(* IEC 61131-3 sources: daoli-st-library/DL_Motion (part 24) *)

(* ---- FB_DL_MotionCmdQueue.st ---- *)
(*
    FB_DL_MotionCmdQueue —— 运动指令排队器（仅 Buffered 语义）
    ------------------------------------------------------------------
    分类      : DL_Motion / CommandMgmt
    前缀      : FB_DL_
    版本      : 1.0.1
    溯源      : T1-6 PLCopen MC_BUFFERMODE 公开条款（Aborting / Buffered / BlendingLow /
                BlendingHigh / BlendingPrevious / BlendingNext 六种，其中 Buffered
                = 「新指令等前一条 Done 之后才影响轴」）；本件只实现 Buffered 一种；
                环形缓冲、满队策略、去重、自愈规则与码位 100% 自有；clean-room 重写，
                未复制任何闭源厂商源码，参考实现仅限 MIT/Apache 许可
    道莅 clean-room 防御性实现：语义借鉴、代码与码位 100% 自有
    平台      : 纯 IEC 61131-3，CODESYS V3.5+ / TwinCAT 3 / InoProShop / Machine Expert 通用
    作者      : 道莅代码库 · PLC编程专家（R22 批 4 · #14）
    ------------------------------------------------------------------
    功能说明  : 把上位连发的定位指令排成先入先出队列，按 Buffered 语义一条一条放给轴：
                前一条轴的 Done 未回就不发下一条。本件不消费轴状态、不发 MC_ 功能块、
                不判断运动是否成功——轴的 Done / Error 由调用方以引脚注入。
    职责边界  : ① 只做 Buffered。Blending 系列不立：BlendingLow / BlendingHigh /
                   BlendingPrevious / BlendingNext 都要求「两段速度在过渡点融合」，
                   而本库的轴侧接口没有速度融合通道，硬做只能做出假混合，
                   比不做更危险——故明确不立项，调用方需融合时请用轴厂家的原生接口。
                ② 不做指令合法性（软限位、速度上限）判定，那是 FB_DL_SoftLimitGuard 的职责。
                ③ bAxisError 到达后只挂起不自动续发：必须先让轴故障消失、再给 bClear，
                   否则队列会在轴仍故障时继续往下砸指令，那是二次伤害。
    队列实现  : 环形缓冲，深度固定 DL_MQ_DEPTH = 8（不参数化：动态内存违反零厂商依赖）。
                头指针指向待发条目，尾指针指向下一个空位，计数 _uCount 为权威值。
    自愈规则  : 每拍前置一致性检查，规则写在此处即此件的契约：
                ① 头指针、尾指针任一 >= DL_MQ_DEPTH，或计数 > DL_MQ_DEPTH
                   → 指针与内容均不可信，整队重建（计数与双指针全部归零）；
                ② 指针均合法时，用 (尾 − 头 + 深度) MOD 深度 反算应有计数，
                   满队时该值为 0，按满队解释为 DL_MQ_DEPTH；
                   反算值与 _uCount 不符 → 以指针为准重建计数（双指针是同拍维护的，
                   计数可能被外部复位或掉电字节残留破坏，指针更可信）。
                自愈是静默的，不占码位（不影响工艺判定），但会在头注释留档供现场排查。
    偏离留档  : 派单写「bAxisDone 上升沿出队」，若按字面在 Done 那一拍才移出队首，
                bClear 期间的槽位归属会与新入队条目混叠（新条目可能被下一次 Done 误当成
                在飞条目弹出，等于吞掉一条指令）。本件把「出队」放在发令那一拍完成，
                Done 只负责把状态机送回 eIdle——语义等价，且消除了混叠路径。
    错误码    : 16#0004_01D9 队列满：bOverwriteOldest=TRUE 丢最旧 / FALSE 拒绝新入队
                              （两策略共用本码，靠 uDropped 是否自增区分）——信息级
                16#0004_01DA 连续同目标同速度的指令已合并去重——信息级，正常防御
                16#0004_02F0 指令参数非有限（NaN / ±Inf），拒绝入队且不占槽——故障级，
                             只拒这一条，不打断整队，也不改变状态机（非锁存）
                16#0004_02F1 轴故障应答（bAxisError），已清队并挂起，禁止自动续发——故障级
                16#0004_02F2 状态机落 ELSE 兜底（非法状态）——故障级，回 eIdle 并清队
    码位总账  : 16#0004_01D9 用 / 16#0004_01DA 用 ｜ 16#0004_02F0 用 / 16#0004_02F1 用 / 16#0004_02F2 用
    状态机    : E_DL_CmdQueueState（eIdle / eSending / eWaitDone / eFault），
                CASE 含 ELSE 兜底，ELSE 置 16#0004_02F2 并回 eIdle 同时清队；
                eSending 是单拍相（发令拍），进相即出相，bExec 因此天然只亮一拍。
    采样约定  : 三个 R_TRIG（入队 / 轴 Done / 轴 Error）在本体最前部无条件刷新（R40）；
                bExec 由段 2 的预置清零保证单拍（R25 三律：置位后本拍即被预置覆盖，
                下一拍必为 FALSE，不存在只置不清）。
    依赖      : 仅 Standard.library（R_TRIG / ABS / MIN / MAX），不引用任何其他 DL_ 子库。
    验收向量  :
                V1 域外早退：fTargetPos = NaN 入队 → 02F0、bError=TRUE、uCount 不变、
                   不占槽，整队继续可用。
                V2 上限截断：连发 9 条 → 第 9 条时 bFull=TRUE；bOverwriteOldest=TRUE
                   → uDropped=1、uCount 仍 8、01D9；置 FALSE → uDropped 不变、01D9、
                   新条目被拒。
                V3 跨段时序：eWaitDone 中 bAxisDone 与下一次 bEnq 同拍 → 本拍先入队
                   （uCount+1）再出相；下一拍才发令，bExec 不连拍。
                V4 恢复首拍：bAxisError 上升沿 → 02F1、清队、eFault；轴故障消失后
                   单独给 bClear → 回 eIdle，队列为空且不发任何残留指令。
    红线自检  : 1 全局变量声明零使用 / 外部变量访问零使用 / 物理地址零使用 —— 通过，全部量经引脚注入
                2 纯 IEC 61131-3 跨平台 —— 通过，仅 Standard.library，无动态内存
                3 防御性编程 —— 通过，数组索引全部前置界检、计数递减前判零、
                   浮点判等用 1.0E-6 容差、非有限值拒绝入队
                4 声明行同行中英双语注释 + 单位 —— 通过，逐行附注（含枚举与数组）
                5 ENUM + CASE 且含 ELSE 兜底 —— 通过
                6 TON / R_TRIG 无条件刷新 —— 通过，段 1 三个沿实例先行调用
                7 无魔法数 —— 通过，深度、容差、计数上限全部 VAR CONSTANT
    修订记录  : 2026-11-16 v1.0.0 首次入库（R22 批 4 · #14）
                2026-11-16 v1.0.1 R22 终审修复：eSending 进相后队列若被 bClear /
                轴故障清空，发令被跳过时改回 eIdle，不再空等永不到来的轴 Done
                （消除「清队竞态 → eWaitDone 挂死」路径，新增 V5 验收向量：
                eIdle 转 eSending 的下一拍给 bClear → 本拍不发令、回 eIdle、bExec 不出现）
*)
TYPE E_DL_CmdQueueState :
(
    eIdle     := 0,      // 空闲，队列非空即进发令相 / idle, a non-empty queue enters the sending phase
    eSending  := 10,     // 单拍发令相，本拍出队并把指令放到执行引脚 / one-scan sending phase, dequeues and publishes the command
    eWaitDone := 20,     // 等轴 Done，未回不发下一条（Buffered 契约）/ waiting for the axis Done, nothing else is issued before it
    eFault    := 30      // 故障，队列已清，需轴故障消失后再给 bClear / fault, the queue is cleared and a bClear is required after the axis fault disappears
);
END_TYPE

FUNCTION_BLOCK FB_DL_MotionCmdQueue
VAR_INPUT
    bEnq             : BOOL;                   // 入队请求，上升沿生效 / enqueue request, effective on the rising edge
    fTargetPos       : REAL;                   // 目标位置 [mm]，非有限即拒收 / target position [mm], a non-finite value is rejected
    fVelocity        : REAL;                   // 运行速度 [mm/s]，非有限即拒收 / travel velocity [mm/s], a non-finite value is rejected
    bAxisDone        : BOOL;                   // 轴 Done 输入，由调用方注入，本件不消费轴状态 / axis Done injected by the caller, no axis state is consumed here
    bAxisError       : BOOL;                   // 轴故障输入，上升沿清队挂起 / axis error input, a rising edge clears the queue and suspends
    bOverwriteOldest : BOOL := TRUE;           // 满队策略：TRUE 丢最旧 / FALSE 拒绝新入队 / full-queue policy, TRUE drops the oldest, FALSE rejects the newcomer
    bClear           : BOOL;                   // 清队电平，为真期间队列保持空且不发令 / clear level, the queue stays empty and nothing is issued while TRUE
END_VAR
VAR_OUTPUT
    bExec            : BOOL;                   // 发令单拍脉冲，只亮一拍 / issue pulse, asserted for exactly one scan
    fExecPos         : REAL;                   // 本拍发出的目标位置 [mm]，保持到下一次发令 / target position issued this scan [mm], held until the next issue
    fExecVel         : REAL;                   // 本拍发出的运行速度 [mm/s]，保持到下一次发令 / travel velocity issued this scan [mm/s], held until the next issue
    uCount           : UINT;                   // 队列内条目数 [条]，0~DL_MQ_DEPTH / number of queued items [pcs], 0~DL_MQ_DEPTH
    bFull            : BOOL;                   // 队列已满 / the queue is full
    uDropped         : UDINT;                  // 累计丢弃条数 [条]，饱和不回绕 / accumulated dropped items [pcs], saturating and never wrapping
    eErr             : UDINT;                  // 错误码，0 表示无错 / error code, 0 means no error
    bError           : BOOL;                   // 故障级标志，仅故障级错误置位 / fault-class flag, set only on fault-level codes
    bValid           : BOOL;                   // 输出可用标志，= NOT bError / outputs valid flag, equals NOT bError
END_VAR
VAR
    fbEnq            : R_TRIG;                 // 入队沿检测实例，无条件刷新 / enqueue edge instance, refreshed unconditionally
    fbDone           : R_TRIG;                 // 轴 Done 沿检测实例，无条件刷新 / axis Done edge instance, refreshed unconditionally
    fbAxisErr        : R_TRIG;                 // 轴故障沿检测实例，无条件刷新 / axis error edge instance, refreshed unconditionally
    _afPos           : ARRAY[0..DL_MQ_DEPTH - 1] OF REAL;   // 队列位置缓存 [mm]，深度与 DL_MQ_DEPTH 同源 / queued positions [mm], depth tied to DL_MQ_DEPTH
    _afVel           : ARRAY[0..DL_MQ_DEPTH - 1] OF REAL;   // 队列速度缓存 [mm/s] / queued velocities [mm/s]
    _uHead           : UINT;                   // 头指针，指向待发条目 / head pointer, points at the next item to issue
    _uTail           : UINT;                   // 尾指针，指向下一个空位 / tail pointer, points at the next free slot
    _uCount          : UINT;                   // 队列条目数（权威值）[条] / item count, the authoritative value [pcs]
    _uExp            : UINT;                   // 由双指针反算的应有计数，自愈用 [条] / count derived from the pointers, used by the self-healing path [pcs]
    _uDroppedAcc     : UDINT;                  // 丢弃计数累加器，饱和不回绕 [条] / dropped accumulator, saturating and never wrapping [pcs]
    _fLastPos        : REAL;                   // 最近一次入队或发令的目标位置，去重用 [mm] / last queued or issued target, used for de-duplication [mm]
    _fLastVel        : REAL;                   // 最近一次入队或发令的速度，去重用 [mm/s] / last queued or issued velocity, used for de-duplication [mm/s]
    _bHaveLast       : BOOL;                   // 去重基准是否已建立 / whether the de-duplication reference exists
    _bParamBad       : BOOL;                   // 本条指令参数非有限标志 / the incoming command carries a non-finite value
    _eState          : E_DL_CmdQueueState;     // 当前状态 / current state
END_VAR
VAR CONSTANT
    DL_MQ_DEPTH      : UINT := 8;              // 队列深度 [条]，固定不参数化 / queue depth [pcs], fixed and never parameterised
    DL_MQ_UDINT_MAX  : UDINT := 16#FFFF_FFFF;  // 丢弃计数饱和上限 [条] / drop-counter saturation bound [pcs]
    DL_MQ_EPS        : REAL := 1.0E-6;         // 去重浮点判等容差 [mm] / de-duplication tolerance [mm]
    DL_MQ_INF_GUARD  : REAL := 4.0E38;         // 非有限幅值判定阈（大于 REAL 最大值）[mm] / non-finite magnitude guard [mm]
END_VAR

// 段 1｜三个沿检测实例无条件周期刷新（红线 6：严禁放入 IF / CASE）
// segment 1, three edge instances refreshed unconditionally
fbEnq(CLK := bEnq);
fbDone(CLK := bAxisDone);
fbAxisErr(CLK := bAxisError);

// 段 2｜输出与错误状态预置（bExec 的单拍性由这里的预置保证，R25 三律）
// segment 2, preset outputs and error status; the preset here is what makes bExec a true one-scan pulse
eErr := 0;                                      // 预置无错误 / preset no error
bError := FALSE;                                // 预置无故障标志 / preset no error flag
bExec := FALSE;                                 // 预置无发令，任何状态想发令必须在本拍重新置位 / preset no issue, any state must assert it again this scan
_bParamBad := FALSE;                            // 预置入队参数合法 / preset the incoming command as legal

// 段 3｜队列自愈：指针越界即整队重建，计数与指针推算不符以指针为准（规则见头注释）
// segment 3, queue self-healing; an out-of-range pointer rebuilds the whole queue and a count mismatch follows the pointers
IF (_uHead >= DL_MQ_DEPTH) OR (_uTail >= DL_MQ_DEPTH) OR (_uCount > DL_MQ_DEPTH) THEN
    _uHead := 0;                                // 指针越界，头归零 / out-of-range head reset
    _uTail := 0;                                // 指针越界，尾归零 / out-of-range tail reset
    _uCount := 0;                               // 内容不可信，计数归零 / untrustworthy content, count reset
    _bHaveLast := FALSE;                        // 去重基准随队一起作废 / the de-duplication reference dies with the queue
ELSE
    _uExp := (_uTail + DL_MQ_DEPTH - _uHead) MOD DL_MQ_DEPTH;   // 由双指针反算应有计数 / derive the count from the pointers
    IF (_uCount > 0) AND (_uExp = 0) THEN
        _uExp := DL_MQ_DEPTH;                   // 满队时头尾重合，按满队解释 / a full queue has coincident pointers, read it as full
    END_IF
    IF _uCount <> _uExp THEN
        _uCount := _uExp;                       // 计数与指针不符，以指针为准重建 / a mismatch follows the pointers, which are maintained every scan
    END_IF
END_IF

// 段 4｜清队电平：只清队列内容，不打断在飞指令的完成等待（Buffered 契约）
// segment 4, the clear level empties the queue but never interrupts the wait of the in-flight command
IF bClear THEN
    _uHead := 0;                                // 头归零 / head reset
    _uTail := 0;                                // 尾归零 / tail reset
    _uCount := 0;                               // 计数归零 / count reset
    _bHaveLast := FALSE;                        // 去重基准作废 / the de-duplication reference is void
END_IF

// 段 5｜轴故障应答：上升沿清队并挂起，绝不自动续发（批 4 统一口径）
// segment 5, axis error response, a rising edge clears the queue and suspends, never resuming automatically
IF fbAxisErr.Q THEN
    _uHead := 0;                                // 头归零 / head reset
    _uTail := 0;                                // 尾归零 / tail reset
    _uCount := 0;                               // 清队，故障后不得留残留指令 / clear the queue, no residual command may survive a fault
    _bHaveLast := FALSE;                        // 去重基准作废 / the de-duplication reference is void
    eErr := 16#0004_02F1;                       // 故障级：轴故障应答已清队并挂起 / fault: the axis error response cleared the queue and suspended
    bError := TRUE;                             // 置故障标志 / raise the fault flag
    _eState := E_DL_CmdQueueState.eFault;       // 挂起，等轴故障消失后再给 bClear / suspend until the axis fault is gone and a bClear arrives
END_IF

// 段 6｜入队处理：参数门禁 → 去重 → 满队策略 → 落槽
// segment 6, enqueue path, parameter gate then de-duplication then the full-queue policy then the slot write
IF fbEnq.Q AND (NOT bClear) AND (_eState <> E_DL_CmdQueueState.eFault) THEN
    // 6.1 参数门禁：非有限一律拒收，不占槽、不动计数
    // parameter gate, a non-finite value is rejected without taking a slot or touching the count
    IF (fTargetPos - fTargetPos) <> (fTargetPos - fTargetPos) THEN
        _bParamBad := TRUE;                     // 目标位置为 NaN / the target position is NaN
    ELSIF ABS(fTargetPos) > DL_MQ_INF_GUARD THEN
        _bParamBad := TRUE;                     // 目标位置为 ±Inf / the target position is infinite
    ELSIF (fVelocity - fVelocity) <> (fVelocity - fVelocity) THEN
        _bParamBad := TRUE;                     // 速度为 NaN / the velocity is NaN
    ELSIF ABS(fVelocity) > DL_MQ_INF_GUARD THEN
        _bParamBad := TRUE;                     // 速度为 ±Inf / the velocity is infinite
    END_IF

    IF _bParamBad THEN
        eErr := 16#0004_02F0;                   // 故障级：指令参数非有限，拒收 / fault: non-finite command parameter, rejected
        bError := TRUE;                         // 只拒这一条，不打断整队 / rejects this item only and never disturbs the rest of the queue
    ELSIF _bHaveLast
          AND (ABS(fTargetPos - _fLastPos) <= DL_MQ_EPS)
          AND (ABS(fVelocity - _fLastVel) <= DL_MQ_EPS) THEN
        eErr := 16#0004_01DA;                   // 信息级：与最近一条同目标同速度，合并去重 / info: identical to the latest command, merged
    ELSIF _uCount >= DL_MQ_DEPTH THEN
        // 6.2 满队：按策略处理，两种策略共用 01D9，靠 uDropped 是否自增区分（R90）
        // full queue, both policies share 01D9 and are told apart by whether uDropped grows
        IF bOverwriteOldest AND (_uCount > 0) THEN
            _uHead := (_uHead + 1) MOD DL_MQ_DEPTH;     // 丢最旧：头前移一格 / drop the oldest by advancing the head
            _uCount := _uCount - 1;                     // 计数先减，随后落槽再加回 / decrement first, the slot write adds it back
            IF _uDroppedAcc < DL_MQ_UDINT_MAX THEN
                _uDroppedAcc := _uDroppedAcc + 1;       // 丢弃计数饱和自增 / saturating increment of the drop counter
            END_IF
            _afPos[_uTail] := fTargetPos;               // 落槽（索引已由指针范围检查保证合法）/ write the slot, the index was validated by the pointer check
            _afVel[_uTail] := fVelocity;                // 落槽速度 / write the queued velocity
            _uTail := (_uTail + 1) MOD DL_MQ_DEPTH;     // 尾前移一格 / advance the tail
            _uCount := _uCount + 1;                     // 计数加回 / add the count back
            _fLastPos := fTargetPos;                    // 更新去重基准位置 / update the de-duplication reference
            _fLastVel := fVelocity;                     // 更新去重基准速度 / update the de-duplication reference
            _bHaveLast := TRUE;                         // 基准已建立 / the reference now exists
            eErr := 16#0004_01D9;                       // 信息级：队列满，已丢最旧 / info: the queue was full and the oldest was dropped
        ELSE
            eErr := 16#0004_01D9;                       // 信息级：队列满，拒绝新入队（uDropped 不变）/ info: full and the newcomer is rejected, uDropped stays
        END_IF
    ELSE
        _afPos[_uTail] := fTargetPos;           // 落槽（索引已由指针范围检查保证合法）/ write the slot, the index was validated by the pointer check
        _afVel[_uTail] := fVelocity;            // 落槽速度 / write the queued velocity
        _uTail := (_uTail + 1) MOD DL_MQ_DEPTH; // 尾前移一格 / advance the tail
        _uCount := _uCount + 1;                 // 计数加一 / increment the count
        _fLastPos := fTargetPos;                // 更新去重基准位置 / update the de-duplication reference
        _fLastVel := fVelocity;                 // 更新去重基准速度 / update the de-duplication reference
        _bHaveLast := TRUE;                     // 基准已建立 / the reference now exists
    END_IF
END_IF

// 段 7｜状态机：eIdle 取队首 → eSending 单拍发令并出队 → eWaitDone 等 Done → eIdle
// segment 7, the state machine, take the head in eIdle, issue and dequeue in the one-scan eSending phase, then wait for Done
CASE _eState OF
E_DL_CmdQueueState.eIdle:
    IF (_uCount > 0) AND (NOT bClear) THEN
        _eState := E_DL_CmdQueueState.eSending;     // 有货且未清队，进发令相 / there is work and no clear, enter the sending phase
    END_IF

E_DL_CmdQueueState.eSending:
    IF (_uCount > 0) AND (_uHead < DL_MQ_DEPTH) THEN
        fExecPos := _afPos[_uHead];                 // 读队首位置（索引前置界检）/ read the head position with a bounds check
        fExecVel := _afVel[_uHead];                 // 读队首速度 / read the head velocity
        bExec := TRUE;                              // 单拍发令，段 2 的预置保证下一拍必为 FALSE / the one-scan issue, the preset guarantees FALSE next scan
        _fLastPos := fExecPos;                      // 去重基准同步为已发条目 / the de-duplication reference follows the issued item
        _fLastVel := fExecVel;                      // 去重基准同步为已发条目 / the de-duplication reference follows the issued item
        _bHaveLast := TRUE;                         // 基准已建立 / the reference now exists
        _uHead := (_uHead + 1) MOD DL_MQ_DEPTH;     // 出队在发令这一拍完成，避免与 bClear 混叠 / dequeue right here so bClear cannot alias the slot
        _uCount := _uCount - 1;                     // 上面的 _uCount > 0 判断已挡住无符号下溢 / the guard above prevents an unsigned underflow
        _eState := E_DL_CmdQueueState.eWaitDone;    // 已真实发令：本相转入等待轴 Done / issued for real, now wait for the axis Done
    ELSE
        _eState := E_DL_CmdQueueState.eIdle;        // 进相后队列被 bClear / 故障清空：无在飞指令，直接回空闲，不得空等永不出现的 Done（R22 终审修复：消除竞态挂死）/ the queue was emptied after entering this phase, no command is in flight, return to idle instead of waiting forever
    END_IF

E_DL_CmdQueueState.eWaitDone:
    IF fbDone.Q THEN
        _eState := E_DL_CmdQueueState.eIdle;        // 前条完成，允许发下一条 / the previous move is done and the next may be issued
    END_IF

E_DL_CmdQueueState.eFault:
    // 退出条件：轴故障已消失且人来清队——两者缺一不可，绝不自动续发
    // exit needs both a vanished axis fault and an operator clear, no automatic resume
    IF bClear AND (NOT bAxisError) AND (NOT fbAxisErr.Q) THEN
        _eState := E_DL_CmdQueueState.eIdle;        // 允许回空闲，队列此时已空；进入故障的这一拍不得退出，否则故障码只闪一拍 / back to idle, but never on the entering scan or the fault code would flash for a single scan
    END_IF

ELSE
    eErr := 16#0004_02F2;                           // 故障级：状态机落 ELSE / fault: the state machine fell into ELSE
    bError := TRUE;                                 // 置故障标志 / raise the fault flag
    _uHead := 0;                                    // 非法态一律清队，绝不带着未知队列继续跑 / an illegal state always clears the queue
    _uTail := 0;
    _uCount := 0;
    _bHaveLast := FALSE;                            // 去重基准作废 / the de-duplication reference is void
    _eState := E_DL_CmdQueueState.eIdle;            // 回空闲 / back to idle
END_CASE

// 段 8｜出口汇总：计数类只做发布，不再二次改写（禁隐式回夹）
// segment 8, exit aggregation; counters are published here and never rewritten again
uCount := _uCount;                              // 队列条目数发布 [条] / publish the queued item count [pcs]
uDropped := _uDroppedAcc;                       // 丢弃累计发布 [条] / publish the accumulated drops [pcs]
bFull := (_uCount >= DL_MQ_DEPTH);              // 满队标志 / full-queue flag
bValid := NOT bError;                           // 输出可用 = 无故障级错误 / outputs are valid when no fault-level code is present
END_FUNCTION_BLOCK

(* ---- FB_DL_PassiveHomingMonitor.st ---- *)
(*==============================================================================
 * 组件名称 (Component)  : FB_DL_PassiveHomingMonitor
 * 所属子库 (Sublibrary) : DL_Motion
 * 当前版本 (Version)    : 1.0.1
 * 组件分类 (Category)   : 功能块（FUNCTION_BLOCK）· 被动回零旁路监听（参考事件确认）
 * 兼容性   (Platform)   : CODESYS 3.5 / TwinCAT 3 / 汇川 InoProShop / Schneider Machine Expert
 *                         仅依赖 Standard.library（R_TRIG / F_TRIG / TON / ABS / MIN / MAX / LIMIT）
 * 接口依赖 (Depends)    : 无 DL_ 内部依赖。本件**不引用**轴状态枚举、**不定义**轴状态枚举，
 *                         也**不调用**任何 MC_ 运动功能块（见分层声明）。
 * 功能描述 (Function)   : 轴被外力移动时（手摇轮、另一驱动拖动、重力下落、维护推车），
 *                         旁路监听参考事件（原点开关沿 / Z 相 / 标记锁存），按「方向一致性
 *                         + 速度窗 + 多次位置一致性」三条判据确认参考点，输出建议施加的
 *                         位置偏移给上层，由上层以 MC_SetPosition 语义消费。
 * 边界（最重要）        : **不自造轴状态、不写轴状态机**。本件只有一个工艺位 bReferenced，
 *                         轴状态（Disabled / Standstill / DiscreteMotion 等）**只由运动层
 *                         拥有**——这是 R31 家族（两套状态机并存）的最高危区，本件按 R11
 *                         判例执行：输出相位 ePhase 仅供 HMI 诊断显示，**不得**被上层当作
 *                         轴状态使用，也不得反向改写轴状态位。
 *                         与 FB_DL_AxisHomingSeq 的分工：后者是**主动回零顺控**（自己发运动
 *                         指令、四模式），本件**不发任何运动指令**，只旁路监听并输出偏移；
 *                         两者可并存，但不得互相改写对方的结论位。
 * 分层声明 (Layer)      : 运动层旁路监视件。上行只为「建议偏移」，下行只有引脚采样。
 *                         零全局变量表引用、零外部变量声明、零物理 IO 地址。
 * 段序     (Segments)   : 段1 实例无条件刷新 → 段2 复位通道（CASE 前，R39）→ 段3 撤防受理 →
 *                         段4 输入防御与镜像量锁定 → 段5 布防受理（倒计置位点，R34）→
 *                         段6 事件受理（倒计递减点，与段5 相邻，R34）→ 段7 状态机 →
 *                         段8 码位单一优先级链 → 段9 出口钳位与保持语义重写。
 * 枚举映射表 (R31)      : eIdle(0)→标签 0｜eArmed(10)→标签 10｜eCaptured(20)→标签 20｜
 *                         eConfirmed(30)→标签 30｜eTimeout(40)→标签 40｜eFault(99)→标签 99。
 *                         每个成员有且仅有一个显式标签，ELSE 只接脏值（02D4）。
 * 单拍标志清单 (R25)    : bArm —— 预清零点：段1 每拍由 `_bArmReq := FALSE` 前的实例输出覆盖；
 *                         置位点：段1 `_bArmReq := _fbTrigArm.Q AND (NOT _bArmConsumed)`；
 *                         自清点：段5 消费时 `_bArmConsumed := TRUE`（撤防、超时、复位三处解除）。
 *                         bReset —— 预清零点：段1 每拍覆盖 _bResetEdge；置位点：段1 的
 *                         _fbTrigReset 实例调用；自清点：紧随实例调用的 _bResetEdge 赋值行。
 *                         bRefEvent —— 内部取上升沿（段1 实例），在段6 单点消费，无对外单拍位。
 * 保持位清单 (R27)      : bReferenced / fRefPos / fOffsetToApply —— 三者逐拍由
 *                         _bRefLatched / _fRefPosHeld / _fOffsetHeld 重写并夹域；
 *                         nEventCount 逐拍由 _nEventCount 转换重写。复位沿清结论。
 * 定时器清单 (R40)      : _fbTonArmTimeout｜IN = (相位 = eArmed 或 eCaptured) AND NOT _bArmBreak｜
 *                         断输入标志 _bArmBreak（每次布防置一拍，本拍 TON 复位 ET）｜
 *                         自清点：段3 无条件 `IF _bArmBreak THEN _bArmBreak := FALSE; END_IF`。
 *                         _fbTonNoMotion｜IN = (相位 = eArmed 或 eCaptured) AND NOT bInMotion
 *                         AND NOT _bArmBreak｜语义为「布防期间长时间静止」信息码 01C5。
 * 三元一致表 (R35)      : 速度窗下限守卫 0.01~100 mm/s / 封顶 100 / 判据 `<`（低于即降精度）｜
 *                         速度窗上限守卫 1~10000 mm/s / 封顶 10000 / 判据 `>`（高于即降精度）｜
 *                         一致性容差守卫 0.001~10 mm / 封顶 10 / 判据 `>`（超出即计数重置）。
 * 镜像量清单 (R38)      : fActPos 的唯一消费点是 _fPosSnap（段4 锁定），fActVel 的唯一消费点
 *                         是 _fVelSnap（段4 锁定）；事件受理与限幅判定全部读快照，不读实时入参。
 * 开源溯源 (Origin)     : 原创实现（参考 PLCopen Part 1 的「参考事件（reference event）」与
 *                         被动回零（passive homing）公开语义，T1-6：参考事件上升沿捕获、
 *                         方向一致性、速度窗内采信、多次事件一致性确认，全部为公开的
 *                         技术概念；实现、状态机、码位与引脚契约 100% 本库独立设计，
 *                         clean-room 编写，未复制任何源码行。许可证说明：PLCopen 规范为
 *                         公开规范条款（非代码），引用其条款语义不构成代码复制风险；
 *                         本文件为本库原创，随本库许可证发布。
 * 验收向量 (Acceptance) :
 *   V1 布防 → 正向 20 mm/s → 两次事件（100.00 / 100.05 mm）→ bReferenced = TRUE、
 *      fRefPos = 100.025（取算术均值，非取首个事件，见设计要点③）。
 *   V2（V-C 方向反转）第二次事件发生在反向 → 16#0004_01C4、计数回到 1、**不得**确认。
 *   V3（V-D 超时恢复）tArmTimeout 到 → eTimeout + 16#0004_02D2；重新 bArm 后计数从 0 重建
 *      （R41：恢复不重头，不允许沿用上次部分计数）。
 *   V4（V-A 非有限）fActVel = NaN → 16#0004_02D3、fRefPos 保持上次确认值（不写脏值）。
 *   V5（R43 出口夹域）撤防后 fOffsetToApply 保持上次值且夹进 ±1.0E6 mm；冷启动首拍输出 0.0。
 * 偏离留档 (Deviation)  :
 *   ① 「目标位置」来源：规格要求输出 fOffsetToApply = 目标 − 参考，但引脚表未给目标值引脚。
 *      本件按「参考事件处应读 0.0 mm」的通用约定输出 fOffsetToApply = 0.0 − fRefPos；若现场
 *      参考点非 0，调用方在消费时叠加其目标值（不新增引脚，避免破坏已冻结的引脚契约）。
 *   ② 速度窗上限的处置：规格给 01C3 的语义是「低于窗下限，采信但精度降级」。高于上限时
 *      定位精度同样不保（可能漏捕获相邻事件），本件并入同一信息码 01C3，语义记为「速度窗
 *      越界，已采信但精度降级」，不新增码位（码位表以规格为准）。
 *   ③ fVelMin > fVelMax 时按对调修复并保持静默（无对应码位），属参数自愈，不改变判定逻辑。
 * 修订历史 (Revision)   :
 *   2026-11-15  v1.0.0  首版入库（Round 13 · 泳道 C · DL_Motion 第 18 件，补 R8 留扩产项）
 *   2026-11-16  v1.0.1  终审修复：段6 事件受理条件补串 bEnable 与 NOT _bFaultCond ——
 *                       原实现下，非有限值检出当拍若恰有参考事件沿，零化快照会被采信，
 *                       极端情形把 0.0 锁存为参考点（坏值穿透到 bReferenced 保持位）
 *============================================================================*)

(*-----------------------------------------------------------------------------
 * 枚举: E_DL_PassiveHomePhase（归属 FB_DL_PassiveHomingMonitor，同文件发布）
 * 用途: 仅内部相位与 HMI 诊断显示，**不是**轴状态，禁止被上层当作轴状态使用。
 *----------------------------------------------------------------------------*)
TYPE E_DL_PassiveHomePhase :
(
    eIdle      := 0,    // 空闲：未布防 / Idle, not armed
    eArmed     := 10,   // 已布防：等待首个参考事件 / Armed, awaiting the first reference event
    eCaptured  := 20,   // 已捕获：事件数未达标，等待后续一致性事件 / Captured, awaiting consistent events
    eConfirmed := 30,   // 已确认：参考点成立，结论保持 / Confirmed, reference established and held
    eTimeout   := 40,   // 超时：布防期内未捕获足够事件 / Timeout, not enough events while armed
    eFault     := 99    // 故障：位置或速度非有限 / Fault, non-finite position or velocity
) UINT;
END_TYPE

FUNCTION_BLOCK FB_DL_PassiveHomingMonitor
VAR_INPUT
    bEnable          : BOOL;                // 使能（Enable），FALSE = 冻结监听并清布防；复位通道不受其屏蔽 / Enable, FALSE stops monitoring
    bReset           : BOOL;                // 复位（Reset），上升沿清结论与锁存 / Rising edge clears the verdict and latches
    bArm             : BOOL;                // 布防（Arm），上升沿开始监听，下降沿撤防 / Rising edge arms, falling edge disarms
    bRefEvent        : BOOL;                // 参考事件电平（Raw reference event），内部取上升沿 / Raw reference event, edge detected inside
    bDirForward      : BOOL := TRUE;        // 本拍运动方向（Current direction），TRUE = 正向，默认 TRUE / TRUE forward, FALSE reverse
    fActPos          : REAL;                // 实际位置（Actual position）[mm]，只读采样，域 −1E7~1E7 / Actual position [mm], read-only
    fActVel          : REAL;                // 实际速度（Actual velocity）[mm/s]，只读采样，域 −1E5~1E5 / Actual velocity [mm/s], read-only
    bInMotion        : BOOL;                // 轴在运动（Axis in motion），速度超噪声带为 TRUE / TRUE when the axis exceeds the noise band
    fVelMin          : REAL := 1.0;         // 速度窗下限（Velocity window low）[mm/s]，域 0.01~100，默认 1.0 / Velocity window low [mm/s]
    fVelMax          : REAL := 500.0;       // 速度窗上限（Velocity window high）[mm/s]，域 1~10000，默认 500.0 / Velocity window high [mm/s]
    nRequireEvents   : INT := 2;            // 需一致性确认的事件次数（Required consistent events）[次]，域 1~3，默认 2 / Required consistent events, 1 to 3
    fConsistencyTol  : REAL := 0.1;         // 事件位置一致性容差（Consistency tolerance）[mm]，域 0.001~10 / Consistency tolerance [mm]
    tArmTimeout      : TIME := T#120S;      // 布防总超时（Arming timeout），域 1 s~1 h，默认 120 s / Arming timeout, default 120 s
END_VAR

VAR_OUTPUT
    bReferenced      : BOOL;                // 参考点已确认（Referenced），保持语义（R27）/ Referenced, held until reset
    fRefPos          : REAL;                // 确认的参考点位置（Confirmed reference position）[mm]，保持语义 / Confirmed reference position [mm], held
    fOffsetToApply   : REAL;                // 建议施加的位置偏移（Offset to apply）[mm]，= 0.0 − fRefPos，夹进 ±1.0E6 / Offset to apply [mm], clamped
    nEventCount      : UINT;                // 本轮布防内已捕获事件数（Events captured in this arming）[次] / Events captured in this arming
    ePhase           : E_DL_PassiveHomePhase;   // 内部相位（Internal phase），**仅供诊断显示** / Internal phase, diagnostics only
    eHealth          : E_DL_Ne107Status;    // 健康态（NE107 health），引用属主 A1 的枚举 / NE107 health, owned by A1
    uDiagCode        : UDINT;               // 诊断码（Diagnostic code），本拍单一优先级链输出 / Diagnostic code, single priority chain
    uErrorId         : UDINT;               // 故障码（Error code），仅故障级码，0 = 无故障 / Fault-level code, 0 = no fault
    bError           : BOOL;                // 故障标志（Error），仅故障级码置位 / TRUE only for fault-level codes
END_VAR

VAR
    _ePhase          : E_DL_PassiveHomePhase := E_DL_PassiveHomePhase.eIdle; // 内部相位（Internal phase）/ Internal phase value
    _bArmReq         : BOOL;                // 布防单拍请求（Arm one-shot request）/ Arm one-shot request
    _bArmConsumed    : BOOL;                // 布防已消费（Arm consumed flag）/ Arm consumed flag
    _bArmBreak       : BOOL;                // 布防段断输入拍（Arm segment input break）/ One-scan break for the arming timers
    _bResetEdge      : BOOL;                // 复位沿单拍标志（Reset one-shot flag）/ Reset one-shot flag
    _bFaultCond      : BOOL;                // 故障条件（Fault condition）/ Fault condition flag
    _uFaultCode      : UDINT;               // 本拍故障级码（Fault-level code this scan）/ Fault-level code of this scan
    _uFaultLatched   : UDINT;               // 故障码锁存（Latched fault code），仅复位沿清除 / Latched fault code, reset only
    _uInfoCode       : UDINT;               // 本拍信息级码（Info-level code this scan）/ Info-level code of this scan
    _fPosSnap        : REAL;                // 位置快照（Position snapshot）[mm]，镜像量唯一消费点入口 / Position snapshot [mm]
    _fVelSnap        : REAL;                // 速度快照（Velocity snapshot）[mm/s]，镜像量唯一消费点入口 / Velocity snapshot [mm/s]
    _fVelAbs         : REAL;                // 速度绝对值（Absolute velocity）[mm/s] / Absolute velocity [mm/s]
    _fVelMinEff      : REAL;                // 生效速度窗下限（Effective window low）[mm/s] / Effective velocity window low [mm/s]
    _fVelMaxEff      : REAL;                // 生效速度窗上限（Effective window high）[mm/s] / Effective velocity window high [mm/s]
    _fConsTolEff     : REAL;                // 生效一致性容差（Effective consistency tolerance）[mm] / Effective consistency tolerance [mm]
    _nReqEff         : INT;                 // 生效事件次数（Effective required events）[次]，钳位 1~3 / Effective required events, clamped 1 to 3
    _nRequireRemain  : INT;                 // 剩余需确认事件数（Remaining events to confirm）[次]，倒计型（R34）/ Remaining events, countdown type (R34)
    _nEventCount     : INT;                 // 本轮已捕获事件数（Events captured this arming）[次] / Events captured this arming
    _fRefSum         : REAL;                // 事件位置累加（Sum of captured positions）[mm] / Sum of captured positions [mm]
    _fRefMean        : REAL;                // 事件位置均值（Mean of captured positions）[mm] / Mean of captured positions [mm]
    _bDirKnown       : BOOL;                // 方向已记录（Direction recorded）/ Direction recorded flag
    _bLastDir        : BOOL;                // 上一次事件方向（Last event direction）/ Direction of the last captured event
    _bRefLatched     : BOOL;                // 参考点锁存（Reference latch），仅复位沿清除 / Reference latch, reset only
    _fRefPosHeld     : REAL;                // 保持的参考位置（Held reference position）[mm] / Held reference position [mm]
    _fOffsetHeld     : REAL;                // 保持的偏移（Held offset）[mm] / Held offset [mm]
    _fbTrigArm       : R_TRIG;              // 布防上升沿（Arm rising edge）/ Arm rising edge detector
    _fbTrigArmFall   : F_TRIG;              // 撤防下降沿（Arm falling edge）/ Arm falling edge detector
    _fbTrigRefEvt    : R_TRIG;              // 参考事件上升沿（Reference event rising edge）/ Reference event rising edge
    _fbTrigReset     : R_TRIG;              // 复位上升沿（Reset rising edge）/ Reset rising edge detector
    _fbTonArmTimeout : TON;                 // 布防总超时（Arming timeout）/ Arming timeout timer
    _fbTonNoMotion   : TON;                 // 静止监视（No-motion watch）/ No-motion watch timer
END_VAR

VAR CONSTANT
    DL_PHM_REAL_MAX  : REAL := 3.4E38;      // 单精度有限值判据幅值（Finite magnitude bound）/ Finite bound for REAL inputs
    DL_PHM_EPS       : REAL := 1.0E-6;      // 浮点防零容差（Divide-guard epsilon）/ Float divide-guard epsilon
    DL_PHM_POS_MAX   : REAL := 1.0E7;       // 位置输入域（Position input bound）[mm] / Position input bound [mm]
    DL_PHM_VEL_MAX   : REAL := 1.0E5;       // 速度输入域（Velocity input bound）[mm/s] / Velocity input bound [mm/s]
    DL_PHM_VMIN_LO   : REAL := 0.01;        // 速度窗下限的下限（Window low lower clamp）[mm/s] / Lower clamp of the window low [mm/s]
    DL_PHM_VMIN_HI   : REAL := 100.0;       // 速度窗下限的上限（Window low upper clamp）[mm/s] / Upper clamp of the window low [mm/s]
    DL_PHM_VMAX_LO   : REAL := 1.0;         // 速度窗上限的下限（Window high lower clamp）[mm/s] / Lower clamp of the window high [mm/s]
    DL_PHM_VMAX_HI   : REAL := 10000.0;     // 速度窗上限的上限（Window high upper clamp）[mm/s] / Upper clamp of the window high [mm/s]
    DL_PHM_TOL_LO    : REAL := 0.001;       // 一致性容差下限（Tolerance lower clamp）[mm] / Tolerance lower clamp [mm]
    DL_PHM_TOL_HI    : REAL := 10.0;        // 一致性容差上限（Tolerance upper clamp）[mm] / Tolerance upper clamp [mm]
    DL_PHM_OFF_MAX   : REAL := 1.0E6;       // 偏移出口夹域（Offset output clamp）[mm] / Offset output clamp [mm]
    DL_PHM_EVT_MIN   : INT  := 1;           // 最少确认事件数（Minimum required events）[次] / Minimum required events
    DL_PHM_EVT_MAX   : INT  := 3;           // 最多确认事件数（Maximum required events）[次] / Maximum required events
    DL_PHM_EVT_MIN_P : INT  := 1;           // 最小捕获事件数（Minimum captured events）[次] / Minimum captured events
    DL_PHM_ERR_TIMEOUT : UDINT := 16#0004_02D2; // 0004_02D2 布防超时未捕获事件【故障级】/ Arm timeout without event, fault level
    DL_PHM_ERR_NONFIN  : UDINT := 16#0004_02D3; // 0004_02D3 位置或速度非有限【故障级】/ Non-finite position or velocity, fault level
    DL_PHM_ERR_STATE   : UDINT := 16#0004_02D4; // 0004_02D4 非法状态兜底【故障级】/ Illegal state fallback, fault level
    DL_PHM_INFO_VEL    : UDINT := 16#0004_01C3; // 0004_01C3 速度窗越界，事件已采信但精度降级【信息级】/ Velocity window exceeded, low precision, info level
    DL_PHM_INFO_DIR    : UDINT := 16#0004_01C4; // 0004_01C4 方向与上次相反，一致性计数重置【信息级】/ Direction reversed, count reset, info level
    DL_PHM_INFO_NOMOT  : UDINT := 16#0004_01C5; // 0004_01C5 布防期间长时间无运动（未超总超时）【信息级】/ No motion during arming, info level
    DL_PHM_INFO_POS    : UDINT := 16#0004_01C6; // 0004_01C6 多次事件位置超容差，计数重置【信息级】/ Position inconsistent, count reset, info level
    DL_PHM_NOMOT_TIME  : TIME  := T#10S;    // 静止判定时长（No-motion detect time）[ms]，默认 10 s / No-motion detect time, default 10 s
END_VAR

// ============================================================================
// 段 1｜实例无条件周期刷新（R7/0.5：严禁置于 IF / CASE 分支内）
//      Unconditional per-cycle refresh of every instance (R7/0.5)
// ============================================================================
_fbTrigArm(CLK := bArm);                        // 布防上升沿（Arm rising edge）
_bArmReq := _fbTrigArm.Q AND (NOT _bArmConsumed);   // 布防单拍请求（R25 置位点）/ Arm one-shot request
_fbTrigArmFall(CLK := NOT bArm);                // 撤防下降沿（Arm falling edge）
_fbTrigRefEvt(CLK := bRefEvent);                // 参考事件上升沿（Reference event rising edge）
_fbTrigReset(CLK := bReset);                    // 复位上升沿（Reset rising edge）
_bResetEdge := _fbTrigReset.Q;                  // 复位单拍标志紧随实例赋值（R25 自清点）

_fbTonArmTimeout(
    IN := ((_ePhase = E_DL_PassiveHomePhase.eArmed) OR (_ePhase = E_DL_PassiveHomePhase.eCaptured))
          AND (NOT _bArmBreak),                 // 断输入拍串入 IN（R40 合规指纹）/ Segment break folded into IN
    PT := tArmTimeout
);                                              // 布防总超时（Arming timeout）
_fbTonNoMotion(
    IN := ((_ePhase = E_DL_PassiveHomePhase.eArmed) OR (_ePhase = E_DL_PassiveHomePhase.eCaptured))
          AND (NOT bInMotion) AND (NOT _bArmBreak), // 静止且布防中（Stationary while armed）
    PT := DL_PHM_NOMOT_TIME
);                                              // 静止监视（No-motion watch）

// 本拍码与条件预置（每拍重算，杜绝跨拍残留）
// Per-scan preset of codes and conditions, no cross-scan residue
_uFaultCode := _uFaultLatched;                  // 故障码以上拍锁存续用（Carry the latched fault code）
_uInfoCode  := 16#0000_0000;                    // 信息级码预清零（Info code preset to zero）
_bFaultCond := FALSE;                           // 故障条件预清零（Fault condition preset FALSE）

// ============================================================================
// 段 2｜复位通道（R39：置于 CASE 之前，且不被掉使能分支屏蔽）
//      Reset path, before CASE and never masked by the disable branch
// ============================================================================
IF _bResetEdge THEN
    _bRefLatched     := FALSE;                  // 参考点锁存清除（Reference latch cleared）
    _fRefPosHeld     := 0.0;                    // 参考位置保持值清零（Held reference position cleared）
    _fOffsetHeld     := 0.0;                    // 偏移保持值清零（Held offset cleared）
    _nEventCount     := 0;                      // 事件计数清零（Event count cleared）
    _nRequireRemain  := 0;                      // 倒计清零（Countdown cleared）
    _fRefSum         := 0.0;                    // 位置累加清零（Position sum cleared）
    _fRefMean        := 0.0;                    // 位置均值清零（Mean cleared）
    _bDirKnown       := FALSE;                  // 方向记录清除（Direction record cleared）
    _bArmConsumed    := FALSE;                  // 布防消费标志清除（Arm consumed flag cleared）
    _uFaultLatched   := 16#0000_0000;           // 故障码锁存清除（Latched fault code cleared）
    _uFaultCode      := 16#0000_0000;           // 本拍故障码随复位清空，防止段8 重新锁存旧码（Clear this scan code）
    IF _ePhase = E_DL_PassiveHomePhase.eFault THEN
        _ePhase      := E_DL_PassiveHomePhase.eIdle;    // 故障态回空闲（Fault phase back to idle）
        _uFaultCode  := 16#0000_0000;           // 故障码随复位清除（Fault code cleared）
        _bFaultCond  := FALSE;                  // 故障条件随复位清除（Fault condition cleared）
    END_IF
END_IF

// ============================================================================
// 段 3｜撤防受理与断输入拍自清（R40：断输入标志在此无条件复位）
//      Disarm handling plus the unconditional self-clear of the segment break
// ============================================================================
IF _bArmBreak THEN
    _bArmBreak := FALSE;                        // 断输入拍自清（Segment break self-cleared after one scan）
END_IF

IF _fbTrigArmFall.Q THEN
    _bArmConsumed   := FALSE;                   // 撤防允许再次布防（Disarm re-enables arming）
    _nEventCount    := 0;                       // 本轮计数作废（Counts voided）
    _nRequireRemain := 0;                       // 倒计作废（Countdown voided）
    _fRefSum        := 0.0;                     // 累加作废（Sum voided）
    _bDirKnown      := FALSE;                   // 方向记录作废（Direction record voided）
    // 撤防只改「相位显示」，且显式排除故障态与已确认态（R39 合法写法①）
    // Disarm only touches the diagnostic phase and explicitly excludes fault and confirmed
    IF (_ePhase <> E_DL_PassiveHomePhase.eFault) AND (_ePhase <> E_DL_PassiveHomePhase.eConfirmed) THEN
        _ePhase := E_DL_PassiveHomePhase.eIdle; // 回空闲（Back to idle）
    END_IF
END_IF

// ============================================================================
// 段 4｜参数钳位 + 输入防御 + 镜像量锁定（R38：每拍只锁一次，后续只读快照）
//      Parameter clamping, input defense and the single per-scan snapshot (R38)
// ============================================================================
_fVelMinEff  := LIMIT(DL_PHM_VMIN_LO, fVelMin, DL_PHM_VMIN_HI);      // 速度窗下限钳位（Window low clamped）
_fVelMaxEff  := LIMIT(DL_PHM_VMAX_LO, fVelMax, DL_PHM_VMAX_HI);      // 速度窗上限钳位（Window high clamped）
_fConsTolEff := LIMIT(DL_PHM_TOL_LO, fConsistencyTol, DL_PHM_TOL_HI); // 一致性容差钳位（Tolerance clamped）
_nReqEff     := nRequireEvents;             // 事件次数直取引脚（Required events taken as-is）
IF _nReqEff < DL_PHM_EVT_MIN THEN
    _nReqEff := DL_PHM_EVT_MIN;             // 下限钳位（Lower clamp）
ELSIF _nReqEff > DL_PHM_EVT_MAX THEN
    _nReqEff := DL_PHM_EVT_MAX;             // 上限钳位（Upper clamp）
END_IF
IF _fVelMinEff > _fVelMaxEff THEN
    _fVelAbs     := _fVelMinEff;            // 借道交换（Borrow the scratch variable to swap）
    _fVelMinEff  := _fVelMaxEff;            // 下限取原上限（Low takes the former high）
    _fVelMaxEff  := _fVelAbs;               // 上限取原下限（High takes the former low）
END_IF

// 输入防御：位置/速度必须落在域内且有限（NaN/Inf 自比不等，等价式判据）
// Input defense: position and velocity must be finite and inside the domain
IF (NOT (fActPos >= (-DL_PHM_POS_MAX) AND fActPos <= DL_PHM_POS_MAX))
OR (NOT (fActVel >= (-DL_PHM_VEL_MAX) AND fActVel <= DL_PHM_VEL_MAX)) THEN
    IF bEnable THEN
        _bFaultCond := TRUE;                // 非有限值即故障（Non-finite input is a fault）
        _uFaultCode := DL_PHM_ERR_NONFIN;   // 0004_02D3 位置或速度非有限【故障级】/ Non-finite input, fault level
    END_IF
    _fPosSnap := 0.0;                       // 快照置零，绝不用脏值（Snapshot zeroed, never the dirty value）
    _fVelSnap := 0.0;                       // 快照置零（Velocity snapshot zeroed）
ELSE
    _fPosSnap := fActPos;                   // 位置快照锁定（Position snapshot latched）
    _fVelSnap := fActVel;                   // 速度快照锁定（Velocity snapshot latched）
END_IF
_fVelAbs := ABS(_fVelSnap);                 // 速度绝对值（Absolute velocity from the snapshot）

// ============================================================================
// 段 5｜布防受理（R34 倒计置位点；R41：每次布防计数从 0 重建）
//      Arming acceptance: the countdown is preset here (R34) and rebuilt from zero (R41)
// ============================================================================
IF _bArmReq AND (NOT _bArmConsumed) AND bEnable
AND (_ePhase <> E_DL_PassiveHomePhase.eFault) THEN
    _bArmConsumed   := TRUE;                // 消费布防请求（Arm request consumed, R25 自清点）
    _ePhase         := E_DL_PassiveHomePhase.eArmed;    // 进布防相位（Enter armed phase）
    _nEventCount    := 0;                   // 计数从 0 重建，不沿用上次部分计数（R41）
    _fRefSum        := 0.0;                 // 累加从 0 重建（Sum rebuilt from zero）
    _bDirKnown      := FALSE;               // 方向记录清除（Direction record cleared）
    _nRequireRemain := _nReqEff;            // 倒计置位（R34 置位点，与段6 递减点相邻）
    _bArmBreak      := TRUE;                // 布防首拍断定时器输入一拍（R40）
END_IF

// ============================================================================
// 段 6｜参考事件受理（R34 倒计递减点，紧跟段5；三判据顺序：方向 → 位置一致性 → 采信）
//      Reference event acceptance: direction, position consistency, then capture (R34)
// ============================================================================
IF _fbTrigRefEvt.Q AND bEnable AND (NOT _bFaultCond)
AND ((_ePhase = E_DL_PassiveHomePhase.eArmed) OR (_ePhase = E_DL_PassiveHomePhase.eCaptured)) THEN
// 本拍故障（非有限）或掉使能时拒绝受理事件：快照已被置零，采信会把脏值写进结论锁存（v1.0.1 修复）
// Events are rejected on a faulted or disabled scan: the snapshot is zeroed and must never be captured

    // 6.1 方向一致性：与上次事件方向相反 → 计数重置（本条同时覆盖「反向拖动」场景）
    //     Direction consistency: a reversal resets the count
    IF _bDirKnown AND (bDirForward <> _bLastDir) THEN
        _uInfoCode      := DL_PHM_INFO_DIR;     // 0004_01C4 方向反转计数重置【信息级】/ Direction reversed, info level
        _nEventCount    := 0;                   // 计数重置（Count reset）
        _fRefSum        := 0.0;                 // 累加重置（Sum reset）
        _nRequireRemain := _nReqEff;            // 倒计重装（Countdown reloaded）
    END_IF

    // 6.2 位置一致性：与已捕获事件的均值偏差超容差 → 计数重置，本次作为首个新事件
    //     Position consistency: a deviation beyond tolerance restarts the count
    IF (_nEventCount >= DL_PHM_EVT_MIN_P) AND (ABS(_fPosSnap - _fRefMean) > _fConsTolEff) THEN
        _uInfoCode      := DL_PHM_INFO_POS;     // 0004_01C6 位置超容差计数重置【信息级】/ Position inconsistent, info level
        _nEventCount    := 0;                   // 计数重置（Count reset）
        _fRefSum        := 0.0;                 // 累加重置（Sum reset）
        _nRequireRemain := _nReqEff;            // 倒计重装（Countdown reloaded）
    END_IF

    // 6.3 采信本事件（速度窗越界不拒绝，只降精度并置信息码）
    //     Capture this event, the velocity window only degrades the precision
    _fRefSum        := _fRefSum + _fPosSnap;    // 位置累加（Position accumulated）
    _nEventCount    := _nEventCount + 1;        // 事件计数 +1（Event counted）
    _nRequireRemain := _nRequireRemain - 1;     // 倒计递减（R34 递减点，与段5 置位点相邻）
    _bDirKnown      := TRUE;                    // 方向记录建立（Direction recorded）
    _bLastDir       := bDirForward;             // 记住本次方向（Remember this direction）
    IF (_fVelAbs < _fVelMinEff) OR (_fVelAbs > _fVelMaxEff) THEN
        _uInfoCode := DL_PHM_INFO_VEL;          // 0004_01C3 速度窗越界精度降级【信息级】/ Velocity window exceeded, info level
    END_IF

    // 6.4 均值重算与结论仲裁（均值取全部已捕获事件，非取首个，见偏离留档①以外的设计要点）
    //     Recompute the mean over every captured event, then arbitrate the verdict
    IF _nEventCount > 0 THEN
        _fRefMean := _fRefSum / INT_TO_REAL(_nEventCount);  // 事件均值（Mean of captured positions），除零已由计数守卫
    END_IF
    IF _nRequireRemain <= 0 THEN
        _bRefLatched := TRUE;                   // 参考点锁存（Reference latched）
        _fRefPosHeld := _fRefMean;              // 参考位置取均值（Reference position takes the mean）
        _fOffsetHeld := 0.0 - _fRefMean;        // 偏移 = 0.0 − 参考（Offset = 0.0 minus the reference）
        _ePhase      := E_DL_PassiveHomePhase.eConfirmed;   // 进已确认相位（Enter confirmed）
    ELSE
        _ePhase := E_DL_PassiveHomePhase.eCaptured;         // 进已捕获相位（Enter captured）
    END_IF
END_IF

// ============================================================================
// 段 7｜状态机（ENUM + CASE，含 ELSE 非法状态兜底）
//      State machine with an explicit ELSE fallback
// ============================================================================
IF _bFaultCond THEN
    _ePhase := E_DL_PassiveHomePhase.eFault;    // 非有限值优先于状态机（Non-finite input outranks the machine）
END_IF

// 掉使能冻结分支：显式排除故障态（R39 合法写法①），复位通道仍可从故障态退出
// Disable branch explicitly excludes the fault state so the reset path still works
IF (NOT bEnable) AND (_ePhase <> E_DL_PassiveHomePhase.eFault) THEN
    _ePhase      := E_DL_PassiveHomePhase.eIdle;    // 冻结回空闲（Freeze back to idle）
    _bArmConsumed := FALSE;                 // 允许重新布防（Arming re-enabled）
    _nEventCount := 0;                      // 计数作废（Counts voided）
    _nRequireRemain := 0;                   // 倒计作废（Countdown voided）
END_IF

CASE _ePhase OF

    E_DL_PassiveHomePhase.eIdle: // 空闲：布防受理已在段5 完成，本分支只保留标签
        // 布防动作在 CASE 之前完成（R39 前置纪律），此处保留空标签与原因注释（R31）
        // Arming happens before CASE, so this label stays empty with its reason (R31)

    E_DL_PassiveHomePhase.eArmed: // 已布防：等首个事件或超时
        IF _fbTonArmTimeout.Q THEN
            _uFaultCode  := DL_PHM_ERR_TIMEOUT;     // 0004_02D2 布防超时【故障级】/ Arm timeout, fault level
            _bFaultCond  := TRUE;                   // 置故障条件（Raise the fault condition）
            _ePhase      := E_DL_PassiveHomePhase.eTimeout; // 进超时相位（Enter timeout）
            _bArmConsumed := FALSE;                 // 允许重新布防（Arming re-enabled）
            _nRequireRemain := 0;                   // 倒计作废（Countdown voided）
        ELSIF _fbTonNoMotion.Q THEN
            _uInfoCode := DL_PHM_INFO_NOMOT;        // 0004_01C5 布防期间长时间无运动【信息级】/ No motion while armed, info level
        END_IF

    E_DL_PassiveHomePhase.eCaptured: // 已捕获：等后续一致性事件或超时
        IF _fbTonArmTimeout.Q THEN
            _uFaultCode  := DL_PHM_ERR_TIMEOUT;     // 0004_02D2 布防超时【故障级】/ Arm timeout, fault level
            _bFaultCond  := TRUE;                   // 置故障条件（Raise the fault condition）
            _ePhase      := E_DL_PassiveHomePhase.eTimeout; // 进超时相位（Enter timeout）
            _bArmConsumed := FALSE;                 // 允许重新布防（Arming re-enabled）
            _nRequireRemain := 0;                   // 倒计作废（Countdown voided）
        ELSIF _fbTonNoMotion.Q THEN
            _uInfoCode := DL_PHM_INFO_NOMOT;        // 0004_01C5 布防期间长时间无运动【信息级】/ No motion while armed, info level
        END_IF

    E_DL_PassiveHomePhase.eConfirmed: // 已确认：结论逐拍在段9 重写，本分支只保留标签
        // 结论保持由段9 逐拍重写承担（R27），此处保留空标签与原因注释（R31）
        // The held verdict is rewritten in segment 9, so this label stays empty (R31)

    E_DL_PassiveHomePhase.eTimeout: // 超时：等重新布防（段5 受理）或复位
        // 重新布防在段5 受理，复位在段2 受理，此处保留空标签与原因注释（R31/R41）
        // Re-arming is accepted in segment 5 and reset in segment 2 (R31/R41)

    E_DL_PassiveHomePhase.eFault: // 故障：等复位沿（段2）
        // 复位通道位于 CASE 之前，此分支无需动作（R39）
        // The reset path sits before CASE, so no action is needed here (R39)

    ELSE // 兜底：非法状态
        _uFaultCode := DL_PHM_ERR_STATE;        // 0004_02D4 非法状态兜底【故障级】/ Illegal state fallback
        _bFaultCond := TRUE;                    // 置故障条件（Raise the fault condition）
        _ePhase     := E_DL_PassiveHomePhase.eFault;    // 强制回故障态（Force the fault state）
END_CASE

// ============================================================================
// 段 8｜码位单一优先级链（全拍只写一次，信息级不置 bError）
//      Single priority chain for the codes, written once per scan
// ============================================================================
IF _uFaultCode <> 16#0000_0000 THEN
    _uFaultLatched := _uFaultCode;              // 故障码锁存，跨拍保持至复位（Latched until reset）
    uErrorId  := _uFaultCode;                   // 故障级码优先（Fault-level code wins）
    uDiagCode := _uFaultCode;                   // 诊断码同源（Diagnostic code mirrors the fault）
    bError    := TRUE;                          // 故障标志置位（Error flag raised）
ELSIF _uInfoCode <> 16#0000_0000 THEN
    uErrorId  := 16#0000_0000;                  // 信息级不占故障码（Info level leaves the fault code empty）
    uDiagCode := _uInfoCode;                    // 诊断码取信息级码（Diagnostic code takes the info code）
    bError    := FALSE;                         // 信息级不置故障位（Info level never raises the error flag）
ELSE
    uErrorId  := 16#0000_0000;                  // 无码（No code）
    uDiagCode := 16#0000_0000;                  // 无码（No code）
    bError    := FALSE;                         // 无故障（No error）
END_IF

// ============================================================================
// 段 9｜出口钳位与保持语义重写（R27/R43：结论逐拍重写，每条路径一次钳位）
//      Output clamping and held-semantics rewrite (R27/R43)
// ============================================================================
bReferenced    := _bRefLatched;                                             // 参考点保持位逐拍重写（Referenced held, rewritten each scan）
fRefPos        := LIMIT(-DL_PHM_OFF_MAX, _fRefPosHeld, DL_PHM_OFF_MAX);     // 参考位置夹进 ±1.0E6（Reference position clamped）
fOffsetToApply := LIMIT(-DL_PHM_OFF_MAX, _fOffsetHeld, DL_PHM_OFF_MAX);     // 偏移夹进 ±1.0E6（Offset clamped）
nEventCount    := INT_TO_UINT(_nEventCount);                                // 事件计数逐拍重写（Event count rewritten）
ePhase         := _ePhase;                                                  // 相位仅供诊断（Phase for diagnostics only）

// 健康态仲裁（引用属主 A1 的四态语言）
// Health arbitration mapped onto the A1 health language
IF _ePhase = E_DL_PassiveHomePhase.eFault THEN
    eHealth := E_DL_Ne107Status.eFailure;       // 故障：信号不可信（Failure）
ELSIF NOT bEnable THEN
    eHealth := E_DL_Ne107Status.eUnknown;       // 未知：未使能（Unknown）
ELSIF _ePhase = E_DL_PassiveHomePhase.eTimeout THEN
    eHealth := E_DL_Ne107Status.eOutOfSpec;     // 越规：布防未取到参考点（Out of spec）
ELSIF _ePhase = E_DL_PassiveHomePhase.eIdle THEN
    eHealth := E_DL_Ne107Status.eUnknown;       // 未知：未布防（Unknown）
ELSE
    eHealth := E_DL_Ne107Status.eOk;            // 正常：监听中或已确认（OK）
END_IF

END_FUNCTION_BLOCK

(* ---- FB_DL_SoftLimitGuard.st ---- *)
(*==============================================================================
 * 组件名称 (Component)  : FB_DL_SoftLimitGuard
 * 所属子库 (Sublibrary) : DL_Motion
 * 当前版本 (Version)    : 1.0.1
 * 兼容性 (Platform)   : CODESYS 3.5 / TwinCAT 3 / 汇川 InoProShop / Machine Expert
 *                         仅依赖 Standard.library（R_TRIG），零厂商方言
 * 分类     (Category)   : 运动安全功能块（Function Block · 软限位电子围栏预判）
 * 功能简述 (Function)   : 软限位安全电子围栏预判器。根据当前速度与减速度实
 *                         时计算双向制动距离（含扫描/IO/驱动时延项），提前
 *                         拦截超程指令；超程后仅允许反向指令（向内恢复豁免
 *                         语义）。位置/速度经既有 I_DL_MotionAxis 接口引用
 *                         读取（fPosition/fVelocity 属性，R11 留档选定）。
 * 定位声明 (Positioning): 公约 0.13——本块为应用层预判与诊断镜像层，不构成
 *                         ISO 13849 / IEC 62061 认证安全功能；硬限位开关与
 *                         认证安全回路的最终防线在认证安全控制器侧，本块输
 *                         出为建议信号（拦截执行在调用方）。
 * 接口消费 (Consumes)   : I_DL_MotionAxis（既有契约，零修改）：读
 *                         iAxis.fPosition / iAxis.fVelocity。R11 二选一留
 *                         档：既有接口已含 fVelocity 速度属性，故不新增
 *                         fAxisSpeed IN_OUT 引脚（规格备选方案弃用）。
 * 公约遵循 (Convention) : 0.1/R23 周期监视型（无初始化/跟踪同步语义），免首
 *                         扫，无 bInit。
 *                         0.2/R21 bFault 显式排除信息级码；0.5/R7 边沿实例主
 *                         体最前部无条件刷新；0.7/R15 故障级锁存仅复位路径清
 *                         码（且离开越界区才可复位）；0.9 全部 REAL 输入/接
 *                         口读数先做非数自比检测（保持末次有效值）；0.14 除
 *                         法带 ABS 防零分支并置码。
 *                         0.8 故障码段位 16#0004_xxxx（经 DL_Motion
 *                         VERSION.md 码表核对：规格建议 0004_0220/0221 已被
 *                         FB_DL_AxisRelativeMove 占用、0004_0106/0107 已占，
 *                         依公约冲突顺延）：
 *                         【故障级】0004_0240 减速度非法、0004_0241 行程边界
 *                         非法；
 *                         【信息级】0004_0108 时延口径提示（默认值与实际不
 *                         符时建议实测，一次性提示）。
 * 红线自检 (Redline)    : R1 零全局变量表/外部变量引用 ✓｜R2 零物理 IO 地址 ✓
 *                         R3 纯 IEC 61131-3 ✓｜R4 除零防御/非有限值防御/浮点
 *                         容差 ✓
 *                         R5 全变量中英双语同行注释 ✓｜R6 N/A（监视型无主状
 *                         态机，判据为纯派生式）✓
 *                         R7 边沿实例主体最前部无条件刷新 ✓｜R8 全常量化 ✓
 * 设计要点 (Key notes)  : ① 预判公式（S-11 提取点①）：fStopDist = fSpeed ×
 *                           tLatency_s + fSpeed² / (2 × fDecel)；tLatency 显
 *                           式换算秒（TIME_TO_REAL 毫秒口径 /1000，舍入意图
 *                           注释写明）；默认 T#23MS 口径 = 扫描 10 + IO 5 +
 *                           驱动 8 ms 三项来源；
 *                         ② 除零防御：fDecel ≤ 1E-6 或非数 → 故障锁存；
 *                           fSpeed² 项在 fSpeed→0 时自然收敛；
 *                         ③ 方向语义：bInterceptPos 置位期间仅允许负向指令
 *                           （向内恢复豁免），本块输出建议信号不直接阻断指
 *                           令（职责边界：拦截执行在调用方）；
 *                         ④ 预警/拦截两级（v1.0.1 勘误：拦截带 ⊇ 预警带——
 *                           拦截含 fMargin 裕量更早触发（保守安全侧），预警带
 *                           为无裕量理论停止距离带；预警带 ⊆ 拦截带，两带
 *                           重合于 fMargin=0 时）；
 *                         ⑤ 参数防御：fPosLimitPos ≤ fPosLimitNeg → 故障锁
 *                           存；复位前提 = 离开越界区（位置回到界内）。
 * 偏离留档 (Deviation)  : 依 R11 头注释留档，共 1 条：
 *                         ① 码位顺延与速度来源：规格建议 0004_0220/0221 与
 *                           既有 FB_DL_AxisRelativeMove 冲突，顺延为
 *                           0004_0240/0241；速度来源选定既有接口属性
 *                           iAxis.fVelocity（规格备选 fAxisSpeed 引脚弃用）。
 * 开源溯源 (Origin)     : 来源标签 plcopen-motion，T1-6 ◐ 深化（RAW_NOTES_R7
 *                         S-11：PLCopen 软限位/Safety-limited 公开语义——
 *                         制动距离预判含时延项、方向性恢复豁免（提取点①②），
 *                         公开规范资料，仅借鉴语义域；预判实现、码位与引脚
 *                         契约 100% 本库独立设计，clean-room 未复制源码）。
 * 验收向量 (Acceptance) :
 *   V1 数值复算：fSpeed=100 mm/s、fDecel=500 mm/s²、tLatency=23MS → 停止距
 *      离 = 100×0.023 + 100²/1000 = 12.3 mm；
 *   V2 预警带进入/退出：位置进入 [边界−停止距离, 边界] → bWarnPos 置位，退
 *      出回落；
 *   V3 双向拦截边界：位置 + 停止距离 + 裕量越界 → bInterceptPos/Neg 置位；
 *   V4 反向恢复豁免：bInterceptPos 期间仅负向指令允许（输出建议语义，注释
 *      写明职责边界）；
 *   V5 参数非法：fDecel=0 → 0004_0240；fPosLimitPos ≤ fPosLimitNeg →
 *      0004_0241；
 *   V6 使能切断仅监视：bEnable=FALSE → 预警照常输出、拦截输出强制 FALSE。
 * 修订历史 (Revision)   :
 *   2026-11-15  v1.0.0  首版入库（Round 07 · DL_Motion 软限位预判件）
 *   2026-11-15  v1.0.1  终审修复 2 处：① fMargin 缺 0.9 非数防御（NaN 时拦
 *                       截比较式恒 FALSE 静默失效），新增 _fMarginEff 生效值
 *                       并钳制负裕量；② 设计要点④「预警带 ⊇ 拦截带」与实
 *                       现/规格向量矛盾，勘误为「拦截带 ⊇ 预警带（含裕量更
 *                       早触发，保守安全侧）」
 *============================================================================*)
FUNCTION_BLOCK FB_DL_SoftLimitGuard
VAR_INPUT
    fPosLimitPos : REAL;                // 正向行程边界（Positive travel limit）[mm]，域 > fPosLimitNeg / Positive travel limit [mm]
    fPosLimitNeg : REAL;                // 负向行程边界（Negative travel limit）[mm] / Negative travel limit [mm]
    fDecel       : REAL := 500.0;       // 拦截减速度（Guard deceleration）[mm/s²]，域 >0，默认 500.0；按配置减速取保守值 / Guard deceleration [mm/s²], conservative value
    tLatency     : TIME := T#23MS;      // 系统-驱动总时延（System latency），默认 T#23MS（扫描 10 + IO 5 + 驱动 8 ms 口径）/ Total latency, default 23 MS (scan 10 + IO 5 + drive 8 ms)
    fMargin      : REAL := 0.0;         // 安全裕量（Safety margin）[mm]，默认 0=关闭裕量；建议 = 停止距离 × 25% / Safety margin [mm], 0 = disabled, suggest 25% of stop distance
    bEnable      : BOOL;                // 预判使能（Guard enable），FALSE=仅监视输出不拦截 / FALSE = monitor only, no intercept
    bReset       : BOOL;                // 上升沿复位故障（Reset edge），离开越界区并复位后方可恢复 / Reset edge, effective only after leaving the overtravel zone
END_VAR
VAR_OUTPUT
    bWarnPos      : BOOL;               // 正向预警（Positive warning），进入「边界 − 停止距离」预判带即置位 / Positive warning inside the limit-minus-stopdist band
    bWarnNeg      : BOOL;               // 负向预警（Negative warning），正向判据镜像 / Mirror of the positive verdict
    bInterceptPos : BOOL;               // 正向拦截（Positive intercept），位置 + 预判停止距离越过边界（含裕量）即置位：调用方应禁止正向指令并减速 / Positive intercept verdict
    bInterceptNeg : BOOL;               // 负向拦截（Negative intercept），正向判据镜像 / Mirror of the positive verdict
    bInsideOk     : BOOL;               // 双向行程内正常（Inside envelope）/ Inside envelope verdict
    fStopDistPos  : REAL;               // 实时正向预判停止距离（Predicted positive stop distance）[mm]，调试/HMI 用 / Predicted stop distance [mm] for HMI
    fStopDistNeg  : REAL;               // 实时负向预判停止距离（Predicted negative stop distance）[mm]，调试/HMI 用 / Predicted stop distance [mm] for HMI
    bFault        : BOOL;               // 故障标志（Fault flag），显式排除信息级 / Fault flag, info codes excluded
    uErrorId      : UDINT;              // 故障码（Error code），16#0004_xxxx 段，0=无故障 / Error code, family 16#0004_xxxx
END_VAR
VAR_IN_OUT
    iAxis        : I_DL_MotionAxis;     // 轴接口引用（Axis interface），由上层注入（既有契约 I_DL_MotionAxis）/ Axis interface reference injected by caller
END_VAR
VAR
    _bFaultLatch  : BOOL;               // 故障锁存标志（Fault latch flag），仅复位路径清除 / Fault latch, cleared only via reset path
    _uErrorIdInt  : UDINT;              // 内部故障级码寄存（Internal fault-level register）/ Internal fault-level register
    _uInfoCode    : UDINT;              // 本拍信息级码（Info code this cycle），瞬时型每拍重算 / Transient info code, recomputed each scan
    _bLatencyHint : BOOL;               // 时延口径提示已发（Latency hint issued）一次性 / One-shot latency hint flag
    _fPosHold     : REAL;               // 末次有效位置保持（Last valid position hold）[mm] / Last valid position hold [mm]
    _fSpdHold     : REAL;               // 末次有效速度保持（Last valid velocity hold）[mm/s] / Last valid velocity hold [mm/s]
    _fPosNow      : REAL;               // 防御后生效位置（Sanitized position）[mm] / Sanitized position [mm]
    _fSpdNow      : REAL;               // 防御后生效速度绝对值（Sanitized speed magnitude）[mm/s] / Sanitized speed magnitude [mm/s]
    _fDecelEff    : REAL := 500.0;      // 防御后生效减速度（Sanitized deceleration）[mm/s²] / Sanitized deceleration [mm/s²]
    _fMarginEff   : REAL;               // 防御后生效安全裕量（Sanitized safety margin）[mm]，0.9 非数防御 / Sanitized safety margin [mm] (v1.0.1)
    _fLatencySec  : REAL;               // 时延秒数（Latency in seconds），TIME 显式换算 / Latency seconds, explicit conversion
    _fStopDist    : REAL;               // 预判停止距离（Predicted stop distance）[mm] / Predicted stop distance [mm]
    _fbTrigReset  : R_TRIG;             // 复位沿（Reset edge）/ Reset edge detector
END_VAR
VAR CONSTANT
    DL_REAL_EPS      : REAL := 1.0E-6;  // 浮点防零容差（Float divide-guard epsilon）/ Float divide-guard epsilon
    DL_TIME_MS_SCALE : REAL := 1000.0;  // TIME→REAL 毫秒换算秒的标度（ms-to-seconds scale）/ Milliseconds-to-seconds scale
END_VAR

// ============================================================================
// 段 1｜实例无条件周期刷新（R7/0.5：严禁置于 IF/CASE 分支内）
//      Unconditional per-cycle refresh of instances (R7/0.5)
// ============================================================================
_fbTrigReset(CLK := bReset);

// ============================================================================
// 段 2｜信息级预清零 + 参数防御（0.9：非数自比，默认值先行）+ 复位路径（R15）
//      Info preset + parameter sanitation (0.9) + reset path (R15)
// ============================================================================
_uInfoCode := 0;                  // 信息级瞬时型每拍重算（Transient info recomputed each scan）

IF fDecel <> fDecel THEN          // 减速度非数自比（Decel NaN self-compare）
    _bFaultLatch := TRUE;         // 减速度非法锁存（Invalid decel latch）
    _uErrorIdInt := 16#0004_0240; // 0004_0240 减速度非法【故障级】/ Invalid deceleration, fault level
ELSIF ABS(fDecel) <= DL_REAL_EPS THEN
    _bFaultLatch := TRUE;         // 减速度趋零防除零锁存（Near-zero decel latch）
    _uErrorIdInt := 16#0004_0240; // 0004_0240 减速度非法【故障级】/ Invalid deceleration, fault level
ELSE
    _fDecelEff := ABS(fDecel);    // 生效减速度（取绝对值保守口径）/ Effective deceleration, magnitude
END_IF

IF fPosLimitPos <= fPosLimitNeg THEN
    _bFaultLatch := TRUE;         // 行程边界非法锁存（Invalid travel limits latch）
    _uErrorIdInt := 16#0004_0241; // 0004_0241 行程边界非法【故障级】/ Invalid travel limits, fault level
END_IF

IF tLatency = T#23MS THEN         // 时延等于默认口径：提示实测（默认值与实际不符建议）
    IF NOT _bLatencyHint THEN
        _bLatencyHint := TRUE;    // 一次性提示标志（One-shot hint flag）
        _uInfoCode := 16#0004_0108; // 0004_0108 时延口径提示【信息级】（建议实测后整定）/ Latency default hint, info level
    END_IF
END_IF
_fLatencySec := TIME_TO_REAL(tLatency) / DL_TIME_MS_SCALE; // TIME→REAL 毫秒口径换算秒（整毫秒时延换算无舍入损失，意图注释）/ ms-to-seconds conversion, exact for whole ms

// 0.9 非数防御补齐（v1.0.1）：fMargin 非数时比较式恒 FALSE → 拦截静默失效
// （安全相关静默降级），非数回落零裕量
// 0.9 NaN defense added (v1.0.1): NaN margin silently disables the intercept
IF fMargin <> fMargin THEN        // 裕量非数（Margin NaN self-compare）
    _fMarginEff := 0.0;           // 回落零裕量（保守域仍由停止距离承担）/ Fallback zero margin
ELSIF fMargin < 0.0 THEN
    _fMarginEff := 0.0;           // 负裕量钳零（防拦截滞后）/ Negative margin clamped to zero
ELSE
    _fMarginEff := fMargin;       // 生效裕量（Effective margin）
END_IF

IF _fbTrigReset.Q AND _bFaultLatch THEN
    // 复位联锁：离开越界区（位置回到界内）且故障源消失才解除
    // Reset interlock: effective only after leaving the overtravel zone
    IF (_fPosHold < fPosLimitPos) AND (_fPosHold > fPosLimitNeg)
       AND (ABS(fDecel) > DL_REAL_EPS) AND (fPosLimitPos > fPosLimitNeg) THEN
        _bFaultLatch := FALSE;    // 故障锁存解除（Fault latch released）
        _uErrorIdInt := 16#0000_0000; // 故障码清零（Fault code cleared）
    END_IF
END_IF

// ============================================================================
// 段 3｜接口读数防御（0.9：非数保持末次有效值）+ 停止距离预判（含时延项）
//      Interface reading sanitation (0.9) + stop-distance prediction with latency
// ============================================================================
IF iAxis.fPosition <> iAxis.fPosition THEN // 位置非数自比（Position NaN self-compare）
    // 保持末次有效位置（Hold last valid position）
ELSE
    _fPosHold := iAxis.fPosition; // 更新末次有效位置（Update last valid position）
END_IF
IF iAxis.fVelocity <> iAxis.fVelocity THEN // 速度非数自比（Velocity NaN self-compare）
    // 保持末次有效速度（Hold last valid velocity）
ELSE
    _fSpdHold := iAxis.fVelocity; // 更新末次有效速度（Update last valid velocity）
END_IF
_fPosNow := _fPosHold;            // 生效位置镜像（Effective position mirror）
_fSpdNow := ABS(_fSpdHold);       // 生效速度幅值（方向由比较式承载）/ Effective speed magnitude (direction carried by comparisons)

_fStopDist := 0.0;                // 出口默认值先赋（Default outlet first）
IF ABS(_fDecelEff) > DL_REAL_EPS THEN
    // 预判公式：时延项 + 制动项（S-11 提取点①）；fSpeed² 项在速度→0 时自然收敛
    // Prediction: latency term + braking term; braking term converges at zero speed
    _fStopDist := (_fSpdNow * _fLatencySec) + (_fSpdNow * _fSpdNow / (2.0 * _fDecelEff)); // 除数已证明非零（Divisor proven non-zero）
END_IF
fStopDistPos := _fStopDist;       // 正向停止距离出口（Positive stop distance outlet）
fStopDistNeg := _fStopDist;       // 负向停止距离出口（对称裕量口径，对称制动力假设）/ Negative outlet (symmetric deceleration assumption)

// ============================================================================
// 段 4｜预警/拦截判据派生（两级：预警带 ⊇ 拦截带；使能切断仅监视）
//      Warning/intercept derivation (two-level, monitor-only when disabled)
// ============================================================================
bWarnPos := (_fPosNow > (fPosLimitPos - _fStopDist)); // 正向预警：进入边界−停止距离带（Positive warning band）
bWarnNeg := (_fPosNow < (fPosLimitNeg + _fStopDist)); // 负向预警镜像（Negative warning mirror）
bInterceptPos := (_fPosNow + _fStopDist + _fMarginEff) > fPosLimitPos; // 正向拦截：含裕量越界预判（生效裕量，v1.0.1）/ Positive intercept with sanitized margin (v1.0.1)
bInterceptNeg := (_fPosNow - _fStopDist - _fMarginEff) < fPosLimitNeg; // 负向拦截镜像（Negative intercept mirror）
IF (NOT bEnable) OR _bFaultLatch THEN
    bInterceptPos := FALSE;       // 使能切断/故障期仅监视：拦截输出强制 FALSE（Monitor-only assertion）
    bInterceptNeg := FALSE;       // 正向断言镜像（Mirror of the positive assertion）
END_IF
bInsideOk := (NOT bWarnPos) AND (NOT bWarnNeg) AND (NOT _bFaultLatch); // 行程内正常派生（Inside-envelope derived form）

// ============================================================================
// 段 5｜方向语义注释（输出建议信号，拦截执行在调用方）+ bFault/uErrorId 出口
//      Direction semantics note + outlets (R21: bFault excludes info codes)
// ============================================================================
// 方向语义（S-11 提取点②）：bInterceptPos 置位期间仅允许负向指令（向内恢复
// 豁免）；bInterceptNeg 置位期间仅允许正向指令。本块输出为建议信号，不直接
// 阻断轴指令——指令禁止与减速执行在调用方（职责边界）。
// Direction semantics: intercept implies opposite-direction commands only; this
// block issues advisory signals only, the caller enforces command blocking.

bFault := _bFaultLatch;           // 故障级派生式（Fault-level derived form）
IF _bFaultLatch THEN
    uErrorId := _uErrorIdInt;     // 故障级码优先透出（Fault-level priority）
ELSE
    uErrorId := _uInfoCode;       // 无故障时透出本拍信息级码（Transient info code）
END_IF
END_FUNCTION_BLOCK

(* ---- FB_DL_SuperimposedMove.st ---- *)
(*==============================================================================
 * 组件名称 (Component)  : FB_DL_SuperimposedMove
 * 所属子库 (Sublibrary) : DL_Motion
 * 当前版本 (Version)    : 1.0.0
 * 分类     (Category)   : 运动工艺功能块（Function Block · 叠加运动补偿层）
 * 作者     (Author)     : Daoli Library
 * 日期     (Date)       : 2026-11-15
 * 兼容性   (Platform)   : CODESYS 3.5 / TwinCAT 3 / 汇川 InoProShop / Schneider
 *                         Machine Expert；纯 IEC 61131-3（第 3 版）语法，
 *                         仅依赖 Standard.library（TON / F_TRIG），零厂商方言
 * 功能简介 (Function)   : 叠加运动补偿层（MC_MoveSuperimposed 语义）。基础轴
 *                         按既有轨迹运行的同时，叠加一个动态偏移量（视觉纠偏、
 *                         张力微调、飞剪对位等场景）；偏移指令经斜坡限速与幅值
 *                         限幅后得到「偏移实际值」，与基础位置相加输出「合成位置」，
 *                         由上层用合成位置下发轴指令。本块只做叠加律、限幅与
 *                         收敛判据，不触碰轴本体指令、不读写轴状态、不做回原。
 *                         与基础运动正交：基础轴正反向运动期间本块无需知情，
 *                         偏移量仅作为位置域的代数叠加项存在。
 * 职责边界 (Scope)      : ① 不产生任何轴使能/定位/停止指令（轴控归上层或
 *                         既有 FB_DL_SingleAxis 类实现块）；② 不读编码器、不做
 *                         位置闭环（纠偏闭环在视觉/张力环内部完成，本块只执行
 *                         已算好的偏移指令）；③ 不做安全限位判断（软限位预判
 *                         归既有 FB_DL_SoftLimitGuard）。
 * 开源溯源 (Origin)     : 来源标签 plcopen-motion / s7-motion（双源印证）。
 *                         仅参考 PLCopen TC3 公开规范与 S7-1500 Motion Control
 *                         公开手册中叠加运动的「功能分类与参数域」（基础运动与
 *                         叠加偏移正交、偏移斜坡限速、零偏移保持叠加层激活的
 *                         行为定义、幅值/速率限制参数域）；本块的状态机、枚举
 *                         编号、引脚契约、故障码位与斜坡实现 100% 本库独立
 *                         设计，clean-room 实现，未复制任何厂商源码行，不构成
 *                         任何来源的衍生作品。
 * 公约遵循 (Convention) : 0.1/R19 首扫范式退化式（本层无外部跟踪源，故取
 *                         IF (NOT bInit) 唯一判据）；0.2/R21 bError 显式排除
 *                         信息级码；0.5/R7 边沿与定时器实例主体最前部无条件
 *                         刷新；0.7/R15 故障级锁存仅重建路径清码；0.9 非有限值
 *                         自比防御 + 出口默认值先赋；0.14 除法与浮点比较全部
 *                         带 ABS 容差；0.16 阈值全常量化。
 * 红线自检 (Redline)    : 全局隔离 ✓（零全局变量表引用、零外部变量声明、零物理
 *                         地址字面记号）｜命名合规 ✓（b/n/u/f/t/a/st/e/fb/i 前缀
 *                         全覆盖）｜注释完整 ✓（声明行 100% 中英双语同行注释）｜
 *                         OOP 封装 ✓（内部状态全私有，仅引脚出口）｜周期安全 ✓
 *                         （TON / F_TRIG 实例无条件刷新）｜防御编程 ✓（除零守卫、
 *                         浮点容差、ENUM + CASE + ELSE 兜底）｜可移植性 ✓（纯
 *                         IEC 61131-3，零厂商私有库）｜终结符成对 ✓
 * 设计要点 (Key notes)  : ① 斜坡实现：本版将斜坡积分内联实现（每拍步进 =
 *                           maxOffsetSpeed × 任务周期），一次乘加即可完成，避免
 *                          REAL/LREAL 与 TIME 毫秒量化的双重精度损失；算法思想
 *                          与已入库 FB_DL_RateLimiter 同源（单向对称限速），
 *                          独立实现、不调用其实例（规格偏离留档见下）。
 *                         ② 限幅次序：先按 bZeroNow 归零目标，再按 maxOffset
 *                          双向幅值钳位，最后进斜坡；钳位发生时置信息级码，
 *                          斜坡仍继续（现场表现为「削顶平移」，不跳变）。
 *                         ③ 零偏移归零完成判据：偏移目标与实际同时落入容差带后
 *                          还需经过零驻留窗口（TON）才判 bInSync，并把浮点残差
 *                          硬置 0.0，防止 HMI 长期显示 0.000001 的假偏移。
 *                         ④ 冻结语义：bEnable = FALSE 时斜坡停走、偏移实际值
 *                          保持（不归零、不跳变），合成位置继续 = 基础 + 保持值；
 *                          重新使能后斜坡从冻结值继续，不产生阶跃（R19 重建式）。
 *                         ⑤ 故障重建：本块故障为参数级（幅值/周期非法）与状态级
 *                          （非法枚举），按规格以 bEnable 下降沿重建回 eIdle，
 *                          重建时清故障码但保持偏移实际值（不归零、不跳变），
 *                          首扫同步只在实例首次运行执行一次。
 * 偏离留档 (Deviation)  : ① 规格 VAR 段列出 fbSlew : FB_DL_RateLimiter 实例，
 *                         实现改为内联斜坡积分（理由见设计要点①，影响：无外部
 *                         组件依赖，引脚契约与输出语义完全不变）；
 *                         ② 规格 VAR 段 bFirstScan 改名 _bInit（理由：公约 0.1
 *                         统一命名 bInit，影响：无）；
 *                         ③ 规格状态跃迁文案「参数非法或斜坡故障 → eFault」中
 *                         斜坡故障项随内联实现取消，参数非法与非法状态两项保留。
 * 故障码表 (Error codes) :
 *                         16#0004_01A0【信息级】任务周期引脚非法已按 10 ms 兜底
 *                         16#0004_01A1【信息级】偏移指令已按幅值上限限幅
 *                         16#0004_01A2【信息级】偏移指令非有限值已拒绝（保持）
 *                         16#0004_01A3【信息级】不限速直通（限速值 <= 0，一次性提示）
 *                         16#0004_02B0【故障级】偏移幅值上限非法（<= 0 或非有限值）
 *                         16#0004_02B1【故障级】任务周期非法（<= 0 或非有限值）
 *                         16#0004_02B2【故障级】非法状态兜底（枚举越界）
 * 验收向量 (Acceptance) :
 *   V1 斜坡跟随：maxOffsetSpeed = 10 mm/s、周期 10 ms、指令跳变 5 mm
 *      → 每拍偏移实际值 +0.1 mm，50 拍后到位，bInSync 置位；
 *   V2 幅值限幅：maxOffset = 5 mm、指令 8 mm → 偏移实际值封顶 5 mm 且
 *      信息级 0004_01A1（每拍重算，超限期间持续）；
 *   V3 零偏移归零判据：指令回 0 → 偏移按斜坡回落，落入容差带后尚需 T#100MS
 *      零驻留窗口，窗口满才 bInSync 且偏移实际值硬置 0.0；
 *   V4 使能冻结：bEnable 下降 → 偏移实际值保持、bActive FALSE、合成位置
 *      仍 = 基础 + 保持值；重新使能斜坡从保持值继续，无阶跃；
 *   V5 参数非法：maxOffset = 0 → 锁 eFault + 0004_02B0；任务周期 0
 *      → 兜底 10 ms + 0004_01A0（周期非法优先钳位，幅值非法才锁故障）；
 *   V6 运行中途插入强制归零：bZeroNow 置位 → 目标立即为 0，斜坡退偏移，
 *      基础位置跟踪不受影响（正交性验证）。
 * 修订历史 (Revision)   :
 *   2026-11-15  v1.0.0  首版入库（Round 09 · DL_Motion 叠加运动补偿件）
 *============================================================================*)

(*-----------------------------------------------------------------------------
 * 调用示例 (Instance guide)：
 *   VAR fbOverlay : FB_DL_SuperimposedMove; END_VAR
 *   fbOverlay(bEnable := bVisionOk,
 *             fBasePos := fbAxis.fPosition,        // 基础轴实际位置注入
 *             fOffsetCmd := fVisionOffset,         // 视觉纠偏量
 *             fMaxOffset := 5.0,
 *             fMaxOffsetSpeed := 10.0,
 *             fTaskCycle := 0.01);                 // 与任务周期一致
 *   fbAxis.MoveAbsolute(fPos := fbOverlay.fSuperPos);  // 用合成位置下发
 *   注意：本块每拍都必须调用（斜坡为逐拍积分，跳拍会丢失积分步长）。
 *----------------------------------------------------------------------------*)

(*-----------------------------------------------------------------------------
 * 常见误用与现场提示 (Field notes)：
 *   1 fTaskCycle 必须与真实任务周期一致：填错会直接放大/缩小偏移速度，本块
 *     无法自检真实周期（禁读 CPU 钟，周期由引脚注入）。
 *   2 合成位置用于下发定位指令时，基础轴必须是位置模式且每拍可接受新目标；
 *     若基础轴为速度模式，请由上层把 fSuperPos 转换为位置增量后再下发。
 *   3 bEnable = FALSE 的语义是「冻结」而非「归零」：需要归零请置 bZeroNow
 *     或把 fOffsetCmd 写 0 后等 bInSync。
 *   4 偏移实际值是纯指令推算量，不含机械跟随误差；精度由基础轴跟随能力决定。
 *   5 幅值上限必须小于安全行程半径，本块不做软限位判断，越界风险由调用方
 *     的软限位预判块承担。
 *----------------------------------------------------------------------------*)

(*-----------------------------------------------------------------------------
 * 枚举: E_DL_OverlayState（归属 FB_DL_SuperimposedMove，随本文件发布）
 * 含义: 叠加补偿层离散状态。数值步长 10 留空位，故障态 99 保证排序末位。
 *----------------------------------------------------------------------------*)
{attribute 'strict'}
{attribute 'qualified_only'}
TYPE E_DL_OverlayState :
(
    eIdle   := 0,    // 空闲：未使能或已冻结，偏移实际值保持 / Idle: disabled or frozen, actual offset held
    eActive := 10,   // 叠加生效：斜坡跟踪偏移指令，零偏移时亦保持本态 / Active: ramp tracks the offset command, zero offset stays active
    eFault  := 99    // 故障锁存：参数或状态非法，输出冻结待重建 / Fault latched: illegal parameter or state, outputs frozen until rebuild
) UINT;
END_TYPE

(*==============================================================================
 * 功能块: FB_DL_SuperimposedMove
 * 调用约定: 每个扫描周期无条件调用一次；全部输入为纯引脚，无任何硬件依赖。
 * 无状态泄漏: 状态仅驻留于实例私有成员，可多实例并行（多轴各一实例）。
 *============================================================================*)
FUNCTION_BLOCK FB_DL_SuperimposedMove
VAR_INPUT
    bEnable         : BOOL;             // 叠加层使能（Overlay enable），FALSE = 斜坡冻结、偏移保持 / FALSE freezes the ramp and holds the offset
    fBasePos        : LREAL;            // 基础轴实际位置（Base axis actual position）[mm]，每拍由上层注入 / Injected each scan by the caller
    fOffsetCmd      : LREAL := 0.0;     // 叠加偏移指令（Offset command）[mm]，正负双向 / Bidirectional offset command [mm]
    fMaxOffset      : LREAL := 5.0;     // 偏移幅值限幅（Offset magnitude limit）[mm]，域 > 0 / Must be greater than zero
    fMaxOffsetSpeed : LREAL := 10.0;    // 偏移斜坡限速（Offset ramp speed limit）[mm/s]，0 = 不限速直通 / Zero means unlimited pass-through
    fTaskCycle      : LREAL := 0.01;    // 任务周期（Task cycle time）[s]，斜坡积分步长基准 / Ramp integration step base in seconds
    bZeroNow        : BOOL;             // 强制归零请求（Force offset to zero）[TRUE = 目标置 0 仍走斜坡] / Target forced to zero, ramp still applied
END_VAR
VAR_OUTPUT
    fSuperPos       : LREAL;            // 合成位置（Superimposed position）[mm] = 基础位置 + 偏移实际值 / Base position plus actual offset
    fOffsetAct      : LREAL;            // 偏移实际值（Actual offset）[mm]，经斜坡与限幅后的代数叠加量 / Ramp-limited and clamped algebraic offset
    bActive         : BOOL;             // 叠加生效中（Overlay active），TRUE = 处于 eActive 态 / TRUE while in the active state
    bInSync         : BOOL;             // 偏移已收敛（Offset in sync），零偏移需驻留窗口满 / Zero offset additionally requires the dwell window
    bError          : BOOL;             // 故障保持型（Fault latched），显式排除信息级码 / Latched fault flag, info codes excluded
    uErrorId        : UDINT;            // 故障码（Error code），0 = 无故障，段位 16#0004_xxxx / Error code, zero means no error
END_VAR
VAR
    _eState         : E_DL_OverlayState := E_DL_OverlayState.eIdle; // 主状态机当前状态（Current state machine state）/ Current state machine state
    _bInit          : BOOL;             // 首扫完成标志（First-scan done flag），初值 FALSE 满足公约 0.1 / First-scan done flag, initial FALSE per convention 0.1
    _bFaultLatch    : BOOL;             // 故障锁存（Fault latch），仅使能下降沿重建路径清除 / Fault latch, cleared only by the disable-edge rebuild path
    _uErrorIdInt    : UDINT;            // 故障级码寄存（Fault-level code register），锁存型 / Latched fault-level code register
    _uInfoCode      : UDINT;            // 本拍信息级码（Info code this scan），每拍重算 / Info code recomputed every scan
    _bRateHint      : BOOL;             // 不限速提示已发（Unlimited-speed hint issued），一次性 / One-shot hint that the ramp is bypassed
    _fMaxOffsetEff  : LREAL := 5.0;     // 生效幅值上限（Effective magnitude limit）[mm]，取绝对值 / Effective magnitude limit, absolute value
    _fRateEff       : LREAL := 10.0;    // 生效斜坡速率（Effective ramp speed）[mm/s]，<= 0 表示直通 / Effective ramp speed, zero or less bypasses the ramp
    _fTaskCycleEff  : LREAL := 0.01;    // 生效任务周期（Effective task cycle）[s] / Effective task cycle in seconds
    _fBaseEff       : LREAL;            // 生效基础位置（Effective base position）[mm]，非有限值保持末次有效 / Effective base position, holds last valid value for non-finite input
    _fBaseHold      : LREAL;            // 末次有效基础位置（Last valid base position）[mm] / Last valid base position [mm]
    _fCmdHold       : LREAL;            // 末次有效偏移指令（Last valid offset command）[mm] / Last valid offset command [mm]
    _fTargetEff     : LREAL;            // 生效偏移目标（Effective offset target）[mm]，限幅后 / Effective offset target after clamping [mm]
    _fDelta         : LREAL;            // 目标与实际偏差（Target minus actual）[mm] / Target minus actual deviation [mm]
    _fStepMax       : LREAL;            // 本拍允许最大偏移步进（Max offset step this scan）[mm] / Max offset step allowed this scan [mm]
    _bGateRun       : BOOL;             // 斜坡运行闸门（Ramp run gate），使能且无故障 / Ramp run gate, enabled and fault free
    _bZeroSettled   : BOOL;            // 零偏移稳定（Zero offset settled），目标与实际均入容差带 / Zero offset settled, target and actual inside tolerance
    _fbTonZeroDwell : TON;              // 零偏移驻留定时器（Zero-offset dwell timer），归零完成判据 / Zero offset dwell timer used by the settled verdict
    _fbTrigDisable  : F_TRIG;           // 使能下降沿（Enable falling edge），故障重建路径触发 / Enable falling edge used by the rebuild path
END_VAR
VAR CONSTANT
    DL_FLOAT_EPS   : LREAL := 1.0E-6;   // 浮点容差（Float epsilon）[mm]，替代判等 / Float epsilon replacing equality comparison [mm]
    DL_CYCLE_FALLBACK : LREAL := 0.01;  // 任务周期兜底值（Task cycle fallback）[s]，非法时生效 / Fallback task cycle applied when illegal [s]
    DL_ZERO_DWELL  : TIME := T#100MS;   // 零偏移驻留窗口（Zero offset dwell window），归零完成判据 / Dwell window of the zero offset verdict
END_VAR

// ============================================================================
// 段 1｜输出确定性默认值先赋（公约 0.9：任何早退路径输出均确定）
//      Deterministic defaults assigned first so every early exit is defined
// ============================================================================
bActive   := FALSE;                    // 生效标志预清零（Active flag pre-cleared）
bInSync   := FALSE;                    // 收敛标志预清零（In-sync flag pre-cleared）
_uInfoCode := 0;                       // 信息级码每拍重算（Info code recomputed every scan）

// ============================================================================
// 段 2｜实例无条件周期刷新（公约 0.5 / R7：严禁置于 IF / CASE 分支内）
//      Unconditional per-cycle refresh of the timer and edge instances
// ============================================================================
_fbTrigDisable(CLK := bEnable);        // 使能下降沿检测（Enable falling edge detection），TON 实例在段 7 无条件刷新（the TON instance is refreshed unconditionally in section 7）

// ============================================================================
// 段 3｜首扫同步（R19 范式退化式：本层无外部跟踪源，仅首扫判据）
//      First-scan synchronization (degraded R19 form, no external track source)
// ============================================================================
IF NOT _bInit THEN
    fOffsetAct  := 0.0;                // 偏移实际值上电从零起步（Offset starts at zero）
    _fBaseHold  := 0.0;                // 基础位置历史清零（Base position history cleared）
    _fCmdHold   := 0.0;                // 偏移指令历史清零（Offset command history cleared）
    _eState     := E_DL_OverlayState.eIdle; // 状态复位为空闲（State reset to idle）
    _bInit      := TRUE;               // 置首扫完成（First-scan done）
END_IF

// ============================================================================
// 段 4｜参数体检与故障锁存（0.16 全常量化；0.2 故障级与信息级分离）
//      Parameter diagnosis with fault latching, fault level split from info level
// ============================================================================
IF (fMaxOffset <> fMaxOffset) OR (ABS(fMaxOffset) <= DL_FLOAT_EPS) THEN
    _bFaultLatch := TRUE;              // 幅值上限非法锁存（Invalid magnitude limit latched）
    _uErrorIdInt := 16#0004_02B0;      // 0004_02B0 偏移幅值上限非法【故障级】（Invalid offset magnitude limit, fault level）
ELSE
    _fMaxOffsetEff := ABS(fMaxOffset); // 生效幅值上限取绝对值（Absolute magnitude limit applied）
END_IF

IF (fTaskCycle <> fTaskCycle) OR (fTaskCycle <= DL_FLOAT_EPS) THEN
    _fTaskCycleEff := DL_CYCLE_FALLBACK; // 周期非法兜底（Illegal cycle falls back）
    _uInfoCode    := 16#0004_01A0;     // 0004_01A0 任务周期非法已兜底【信息级】（Task cycle fell back, info level）
ELSE
    _fTaskCycleEff := fTaskCycle;       // 合法周期直通（Valid cycle passed through）
END_IF

IF fMaxOffsetSpeed <> fMaxOffsetSpeed THEN
    _fRateEff := 0.0;                  // 非有限限速按直通处理（Non-finite speed bypasses the ramp）
ELSIF fMaxOffsetSpeed <= DL_FLOAT_EPS THEN
    _fRateEff := 0.0;                  // 零或负限速按直通处理（Zero or negative speed bypasses the ramp）
    IF NOT _bRateHint THEN
        _bRateHint := TRUE;            // 一次性提示标志（One-shot hint flag）
        _uInfoCode := 16#0004_01A3;    // 0004_01A3 不限速直通提示【信息级】（Ramp bypassed hint, info level）
    END_IF
ELSE
    _fRateEff := fMaxOffsetSpeed;       // 合法限速直通（Valid ramp speed passed through）
END_IF

// ============================================================================
// 段 5｜非有限值防御（0.9：自比检测，保持末次有效值，不中断扫描）
//      Non-finite defense holding the last valid value, scan is never stopped
// ============================================================================
IF fBasePos <> fBasePos THEN
    _fBaseEff := _fBaseHold;           // 基础位置非有限保持末次有效（Non-finite base position holds last valid）
ELSE
    _fBaseHold := fBasePos;             // 更新末次有效基础位置（Last valid base position updated）
    _fBaseEff  := fBasePos;             // 生效基础位置（Effective base position）
END_IF

IF fOffsetCmd <> fOffsetCmd THEN
    _fTargetEff := _fCmdHold;           // 指令非有限保持末次有效目标（Non-finite command holds last valid target）
    _uInfoCode  := 16#0004_01A2;        // 0004_01A2 偏移指令非有限已拒绝【信息级】（Non-finite offset command rejected, info level）
ELSE
    _fCmdHold   := fOffsetCmd;          // 更新末次有效偏移指令（Last valid offset command updated）
    _fTargetEff := fOffsetCmd;          // 生效偏移目标（Effective offset target）
END_IF

// ============================================================================
// 段 6｜目标选取与双向幅值限幅（先归零后限幅，限幅不阻断斜坡）
//      Target selection and symmetric clamping, clamping never blocks the ramp
// ============================================================================
IF bZeroNow THEN
    _fTargetEff := 0.0;                // 强制归零优先（Force-zero takes priority）
END_IF

IF ABS(_fTargetEff) > _fMaxOffsetEff THEN
    IF _fTargetEff > 0.0 THEN
        _fTargetEff := _fMaxOffsetEff; // 正向削顶（Clamped at the positive limit）
    ELSE
        _fTargetEff := -_fMaxOffsetEff; // 负向削顶（Clamped at the negative limit）
    END_IF
    _uInfoCode := 16#0004_01A1;        // 0004_01A1 偏移指令已限幅【信息级】（Offset command clamped, info level）
END_IF

// ============================================================================
// 段 7｜斜坡积分与零偏移归零判据（内联斜坡，每拍一步乘加）
//      Inline ramp integration plus the zero-offset settled verdict
// ============================================================================
_bGateRun := bEnable AND (NOT _bFaultLatch); // 运行闸门（Run gate）

IF _bGateRun THEN
    _fDelta := _fTargetEff - fOffsetAct; // 目标与实际偏差（Target minus actual deviation）
    IF _fRateEff <= DL_FLOAT_EPS THEN
        fOffsetAct := _fTargetEff;     // 不限速直通（Unlimited pass-through）
    ELSE
        _fStepMax := _fRateEff * _fTaskCycleEff; // 本拍允许步进 [mm]（Max step this scan）
        IF ABS(_fDelta) <= _fStepMax THEN
            fOffsetAct := _fTargetEff; // 一步到位，杜绝残差抖动（One-step landing avoids residual jitter）
        ELSIF _fDelta > 0.0 THEN
            fOffsetAct := fOffsetAct + _fStepMax; // 正向推进（Advance in the positive direction）
        ELSE
            fOffsetAct := fOffsetAct - _fStepMax; // 负向推进（Advance in the negative direction）
        END_IF
    END_IF
END_IF

_bZeroSettled := (ABS(_fTargetEff) < DL_FLOAT_EPS) AND (ABS(fOffsetAct) < DL_FLOAT_EPS) AND _bGateRun; // 零偏移稳定判据（Zero offset settled verdict）
_fbTonZeroDwell(IN := _bZeroSettled, PT := DL_ZERO_DWELL); // 驻留窗口计时（Dwell window timing）

IF _fbTonZeroDwell.Q THEN
    fOffsetAct := 0.0;                 // 驻留满后硬置零，消除浮点残差（Hard zero after dwell removes float residual）
END_IF

bInSync := (ABS(_fTargetEff - fOffsetAct) < DL_FLOAT_EPS) AND _bGateRun; // 收敛判据：目标与实际偏差入容差带（Convergence verdict within tolerance）
IF (ABS(_fTargetEff) < DL_FLOAT_EPS) AND (NOT _fbTonZeroDwell.Q) THEN
    bInSync := FALSE;                  // 零偏移需驻留窗口满才算归零完成（Zero offset requires the dwell window）
END_IF

// ============================================================================
// 段 8｜主状态机（ENUM + CASE + ELSE 兜底；故障重建走使能下降沿）
//      Main state machine with mandatory ELSE fallback and disable-edge rebuild
// ============================================================================
CASE _eState OF

    E_DL_OverlayState.eIdle: // 空闲：等待使能（Idle, waiting for enable）
        IF _fbTrigDisable.Q THEN
            _bFaultLatch := FALSE;     // 下降沿重建：清故障锁存（Rebuild clears the fault latch）
            _uErrorIdInt := 16#0000_0000; // 故障码清零（Fault code cleared）
        END_IF
        IF bEnable AND (NOT _bFaultLatch) THEN
            _eState := E_DL_OverlayState.eActive; // 使能且参数合法进叠加态（Enabled and legal, go active）
        END_IF

    E_DL_OverlayState.eActive: // 叠加生效：零偏移亦保持本态（Active, zero offset keeps this state）
        IF _bFaultLatch THEN
            _eState := E_DL_OverlayState.eFault; // 参数或状态故障锁存（Fault latched）
        ELSIF NOT bEnable THEN
            _eState := E_DL_OverlayState.eIdle;  // 禁止使能冻结偏移并回空闲（Disable freezes the offset and returns to idle）
        END_IF

    E_DL_OverlayState.eFault: // 故障锁存：输出冻结为最后安全值（Fault latched, outputs frozen）
        IF _fbTrigDisable.Q THEN
            _bFaultLatch := FALSE;     // 使能下降沿重建（Rebuild on the enable falling edge）
            _uErrorIdInt := 16#0000_0000; // 故障码清零（Fault code cleared）
            _eState := E_DL_OverlayState.eIdle; // 回空闲（Back to idle）
        END_IF

    ELSE
        _bFaultLatch := TRUE;          // 非法状态兜底锁存（Illegal state fallback latched）
        _uErrorIdInt := 16#0004_02B2;  // 0004_02B2 非法状态兜底【故障级】（Illegal state fallback, fault level）
        _eState := E_DL_OverlayState.eFault; // 进故障态（Enter the fault state）
END_CASE

// ============================================================================
// 段 9｜出口映射（合成位置 = 基础 + 偏移；故障级码优先透出）
//      Outlet mapping, fault-level code has priority over info codes
// ============================================================================
fSuperPos := _fBaseEff + fOffsetAct;   // 叠加律：代数相加（Superposition as an algebraic sum）
bActive   := (_eState = E_DL_OverlayState.eActive); // 生效标志派生（Active flag derived from the state）
bError    := _bFaultLatch OR (_eState = E_DL_OverlayState.eFault); // 故障派生，显式排除信息级（Fault derived, info codes excluded）
IF bError THEN
    uErrorId := _uErrorIdInt;          // 故障级码优先（Fault-level code has priority）
ELSE
    uErrorId := _uInfoCode;            // 无故障透出本拍信息级码（Transient info code exposed）
END_IF
END_FUNCTION_BLOCK
